(* IEC 61131-3 sources: daoli-st-library/DL_Process (part 34) *)

(* ---- FB_DL_FirstArticleLock.st ---- *)
(*
  ==================================================================
  组件名 Component  : FB_DL_FirstArticleLock
  分类   Category   : DL_Process
  复杂度 Complexity  : cx5
  版本   Version    : 1.0.0
  功能   Purpose    : 首件检验锁定。首件未放行禁止批量运行（许可出口挂锁定
                      状态量）；换型信号沿自动重锁；首件检验合格沿解锁放行
                      并出单拍放行脉冲与台账；锁定期的运行请求出单拍拒绝
                      指示。汽车 / 电子行业公开首件流程语义。
  来源   Source     : self（行业公开流程）
  溯源   Origin     : IEC 61131-3 标准语义的道莅防御性实现；首件检验锁定为
                      公开行业流程语义，clean-room 自研实现，未复制任何厂商
                      私有库源码。
  平台   Platform   : 纯 IEC 61131-3（Standard.library: R_TRIG，无私有库）
  分工声明 Split     : 与 FB_DL_MaterialHoldTimeEnforce 分工——保持时限件做
                      在制批次时限门控，本件做换型后批量运行前置门控；与
                      存量批次追溯件分工——本件不含履历数据，只有锁存与台账。
  作者   Author     : 道莅代码库 · PLC 编程专家（R58）
  ------------------------------------------------------------------
  边界 Boundary     :
                      一 上电默认锁定（_bInit 首扫置锁）：首件未放行禁止批
                         量运行，安全侧缺省；
                      二 锁定解除路径 = bFaPass 上升沿（唯一解锁路径，R188
                         头注释声明）；重锁路径 = bChangeover 上升沿（换型
                         自动重锁）；
                      三 许可出口挂状态量 _bLocked（R99：禁挂单拍标志）；
                      四 单拍标志 bFaRelease / bRunBlocked 每拍预清零（R25，
                         置位点在段 3，统一出口单拍映射两段式 R189）；
                      五 复位沿作用域：清台账 / 恢复默认锁定（两项逐项声明）；
                      六 无全局变量、无外部变量声明、无物理地址寻址。
  修订记录 Revision  :
    2026-11-21  v1.0.0  R58 首版（批 4 · 序号 16）
  ==================================================================
*)

FUNCTION_BLOCK FB_DL_FirstArticleLock
VAR_INPUT
    bEnable     : BOOL := TRUE;   // 使能，失能许可出口安全侧 FALSE [-] / enable, disabling clears the permit
    bReset      : BOOL := FALSE;  // 复位上升沿清台账并恢复默认锁定 [-] / reset rising edge clears the ledger and restores the default lock
    bChangeover : BOOL := FALSE;  // 换型信号（沿生效，自动重锁）[-] / the changeover signal, edge effective, auto relock
    bFaPass     : BOOL := FALSE;  // 首件检验合格（沿生效）[-] / the first article pass, edge effective
    bRunReq     : BOOL := FALSE;  // 批量运行请求电平 [-] / the batch run request level
END_VAR
VAR_OUTPUT
    bBatchPermit: BOOL := FALSE; // 批量运行许可出口（挂锁定状态量）[-] / the batch run permit outlet, gated by the lock state
    bLocked     : BOOL := FALSE; // 锁定中指示出口 [-] / the locked indicator outlet
    bFaRelease  : BOOL := FALSE; // 首件放行单拍出口 [-] / the first article release pulse outlet
    bRunBlocked : BOOL := FALSE; // 锁定期运行请求拒绝单拍出口 [-] / the run request blocked pulse outlet
    nLockCnt    : UDINT := 0;    // 累计重锁次数 [次] / the total relock count
    nRelCnt     : UDINT := 0;    // 累计放行次数 [次] / the total release count
END_VAR
VAR
    rtChg   : R_TRIG; // 换型沿检测，段 0 无条件刷新 / the changeover edge
    rtPass  : R_TRIG; // 首件合格沿检测，段 0 无条件刷新 / the pass edge
    rtReset : R_TRIG; // 复位沿检测，段 0 无条件刷新 / the reset edge
    _bLocked: BOOL := TRUE;  // 锁定状态量（上电缺省锁定，边界一）/ the lock state, the power up default locked
    _bRel   : BOOL := FALSE; // 放行脉冲内部保持量（统一出口映射单拍）/ the release pulse internal holder
    _bBlk   : BOOL := FALSE; // 拒绝脉冲内部保持量 / the blocked pulse internal holder
    _bInit  : BOOL := FALSE; // 首扫初始化完成标志（R310）/ the first scan flag
END_VAR
VAR CONSTANT
    DL_FAL_CNTMAX : UDINT := 4294967294; // 台账计数钳定界 [次]，防 UDINT 回绕 / the ledger clamp against a wrap
END_VAR

// 段 0｜沿检测无条件周期刷新（禁入分支，FB50-1）/ segment 0, the unconditional refresh
rtChg(CLK := bChangeover); // 换型沿 / the changeover edge
rtPass(CLK := bFaPass); // 合格沿 / the pass edge
rtReset(CLK := bReset); // 复位沿 / the reset edge

// 段 1｜首扫初始化（R310）：上电默认锁定（边界一）/ segment 1, the first scan, the default locked
IF NOT _bInit THEN // 首扫一拍 / the first scan
    _bInit := TRUE; // 置首扫标志 / raise the flag
    _bLocked := TRUE; // 上电默认锁定 / the default locked
END_IF

// 段 2｜复位沿作用域：清台账 / 恢复默认锁定（两项逐项声明，边界五）/ segment 2, the reset edge scope
IF rtReset.Q THEN // 复位沿 / the reset edge
    nLockCnt := 0; // 作用域一：清重锁台账 / scope one, clear the relock ledger
    nRelCnt := 0; // 作用域一：清放行台账 / scope one, clear the release ledger
    _bLocked := TRUE; // 作用域二：恢复默认锁定（安全侧）/ scope two, restore the default lock
END_IF

// 段 3｜重锁与解锁沿判定 + 单拍保持量置位（边界二三四）/ segment 3, the relock and the unlock edges
IF rtChg.Q THEN // 换型沿自动重锁 / the changeover edge relocks
    _bLocked := TRUE; // 置锁定 / raise the lock
    IF nLockCnt < DL_FAL_CNTMAX THEN // 台账防回绕 / the ledger wrap guard
        nLockCnt := nLockCnt + 1; // 重锁台账推进 / advance the relock ledger
    END_IF
END_IF
IF _bLocked AND rtPass.Q THEN // 锁定中且首件合格沿（唯一解锁路径，R188）/ locked with the pass edge
    _bLocked := FALSE; // 解锁 / release the lock
    IF nRelCnt < DL_FAL_CNTMAX THEN // 台账防回绕 / the ledger wrap guard
        nRelCnt := nRelCnt + 1; // 放行台账推进 / advance the release ledger
    END_IF
    _bRel := TRUE; // 置放行内部保持量 / raise the release holder
END_IF
IF _bLocked AND bRunReq THEN // 锁定期收到运行请求 / a run request while locked
    _bBlk := TRUE; // 置拒绝内部保持量 / raise the blocked holder
END_IF
bFaRelease := FALSE; // 放行单拍每拍预清零（R25）/ the release pulse preset false each scan
bRunBlocked := FALSE; // 拒绝单拍每拍预清零（R25）/ the blocked pulse preset false each scan

// 段 4｜统一出口（边界三四：状态量门控 + 单拍两段式映射）/ segment 4, the unified outlet
bBatchPermit := (NOT _bLocked) AND bEnable; // 许可挂锁定状态量（R99）/ the permit gated by the lock state
bLocked := _bLocked; // 锁定指示同源 / the indicator shares the state
IF _bRel THEN // 放行保持量 → 统一出口单拍映射（两段式，R189）/ the holder mapped to the pulse
    bFaRelease := TRUE; // 放行单拍 / the release pulse
    _bRel := FALSE; // 消费保持量 / consume the holder
END_IF
IF _bBlk THEN // 拒绝保持量 → 统一出口单拍映射 / the holder mapped to the pulse
    bRunBlocked := TRUE; // 拒绝单拍 / the blocked pulse
    _bBlk := FALSE; // 消费保持量 / consume the holder
END_IF
END_FUNCTION_BLOCK

(* ---- FB_DL_FloatBathTopRollSeq.st ---- *)
(*
  Name: FB_DL_FloatBathTopRollSeq
  Category: DL_Process
  Version: 1.0.0
  Round: R90 / 2026-11-25
  开源溯源：clean-room 自研（族 浮法玻璃锡槽退火，ST 开源生态实测 0 命中，无外部代码引入）
  功能：1) 拉边机三轴同步作业序，六相推进：待机 → 就位 → 夹持 → 同步张角 → 跟踪带宽 → 退出 → 完成。
           就位相向三轴发出就位指令并等三路到位信号全为 TRUE；夹持相保持指令并等夹持时长；
           同步张角相把张角给定按设定角速度斜坡推到 fAngleTargetDeg；跟踪带宽相保持张角并监视
           带宽是否漂出容差；退出相撤令（三轴回退），等退到位时长后置完成位。
        2) 多轴失步监视贯穿三轴：就位相超时未全部到位 → 失步故障；同步相与跟踪相内任一路到位
           信号掉线 → 失步故障。三轴指令始终同源（同一个状态量导出），不存在单轴独走的可能。
        3) 张角斜坡按「角速度 × 扫描周期」逐拍累加，故扫描周期必须作为入参并做零闸（R21），
           不许假设固定扫描周期；斜坡单向逼近目标，不越过目标值。
  边界条件：1) 非有限值闸：张角目标、带宽实测、扫描周期三路实值入参统一过
           NOT(x > -DL_BIG AND x < DL_BIG)，同时拦 NaN 与 Inf；命中即判组态非法并进故障相，
           绝不把 NaN 累加进张角保持值（累加后保持值被永久污染，R19）。
        2) 组态零闸：ABS(fCycleS) > DL_EPS 才允许角度积分（周期为零则斜坡不推进且步进发散）；
           tSyncS 必须 > T#0S（跟踪相时长为 0 表示跳过跟踪监视，属组态错误）；
           fAngleTargetDeg 必须落在 0 ~ DL_ANGLE_MAX_DEG(90 °) 并大于 0。
        3) 带宽容差闸：跟踪相内带宽相对漂移超过 DL_WIDTH_TOL_PCT(2 %) 判带宽失控故障；
           带宽参考值在进入跟踪相的同一个周期末锁存（R23：快照必须在迁移判断之后更新）。
        4) 相超时说明：eFbtPosition 由 tonPos 监视（就位超时 = 失步）；
           eFbtClamp 由 tonClamp 定时（夹持时长，无额外超时）；
           eFbtSyncAngle 由 tonAngle 监视（张角同步超时 = 失步）；
           eFbtTrackWidth 由 tonTrack 定时（跟踪时长，另有带宽容差监视）；
           eFbtRetract 由 tonRetract 定时（退出时长）；
           eFbtDone / eFbtIdle / eFbtFault 为稳态持留相，不设相超时（设了会周期性误报）；
           整序另设 tonSeq 总超时兜底。
        5) 状态机兜底：CASE 全态覆盖 + ELSE 强制回故障相并撤全部指令；故障解除路径为
           (NOT xStart) AND (NOT xFault) AND 组态恢复，可达。
        6) FB 主体不使用 RETURN，统一单出口（跨平台可移植性）。
  量纲自证：张角步进 = (°/s) × s = °，与 fAngleDeg 同量纲；
           带宽相对漂移 = (mm − mm) / mm × 100 = 无因次 [%]，与容差同量纲；
           三路到位信号为 [bool]；tonXxx 的 PT 均为 [TIME]；本件无跨量纲相加。
  码表 Error codes（本件格 0090_07xx，故障级一律 3 行内置 _uFault/_bFault/_eState）:
    16#0090_0701 故障级：组态非法（角度目标/跟踪时长/扫描周期越界或非有限）
    16#0090_0702 故障级：就位超时（三轴未全部到位，多轴失步）
    16#0090_0703 故障级：张角同步超时（斜坡未在时限内到达目标）
    16#0090_0704 故障级：同步/跟踪相内到位信号掉线（多轴失步）
    16#0090_0705 故障级：跟踪相带宽漂移超容差（带宽失控）
    16#0090_0706 故障级：整序总超时
    16#0090_0707 故障级：外部故障输入 xFault
    16#0090_0708 故障级：状态机落 ELSE 兜底（非法相位 ID）
    16#0090_0709 信息级：张角已到达目标，转入跟踪相

  修订历史 Revision :
    2026-11-25  v1.0.0  R90 首版
*)

TYPE E_DL_FbtState :
(
    eFbtIdle      := 0,    // 待机：等启动上升沿 / Idle, awaiting start edge
    eFbtPosition  := 10,   // 就位：三轴发出就位指令 / Positioning, all three axes commanded
    eFbtClamp     := 20,   // 夹持：保持指令等夹持时长 / Clamping, commands held
    eFbtSyncAngle := 30,   // 同步张角：斜坡推到目标角 / Angle synchronising
    eFbtTrackWidth:= 40,   // 跟踪带宽：保持张角并监视带宽 / Width tracking
    eFbtRetract   := 50,   // 退出：撤令等退到位 / Retracting
    eFbtDone      := 60,   // 完成：保持完成位等撤令 / Done, held until release
    eFbtFault     := 90    // 故障：锁存待解除 / Fault, latched awaiting release
);
END_TYPE

FUNCTION_BLOCK FB_DL_FloatBathTopRollSeq
VAR_INPUT
    xStart          : BOOL;    // 作业启动指令（上升沿有效）[bool] / Sequence start, edge triggered [bool]
    xFault          : BOOL;    // 外部故障汇总 [bool] / External fault aggregate [bool]
    xInPos1         : BOOL;    // 1 轴到位信号 [bool] / Axis 1 in-position signal [bool]
    xInPos2         : BOOL;    // 2 轴到位信号 [bool] / Axis 2 in-position signal [bool]
    xInPos3         : BOOL;    // 3 轴到位信号 [bool] / Axis 3 in-position signal [bool]
    fAngleTargetDeg : REAL;    // 目标张角 [°] / Target nip angle [°]
    fWidthMeasMm    : REAL;    // 玻璃带宽度实测 [mm] / Measured ribbon width [mm]
    tSyncS          : TIME;    // 带宽跟踪监视时长 [TIME] / Width tracking supervision duration [TIME]
    fCycleS         : REAL;    // 扫描周期 [s] / Scan cycle time [s]
END_VAR
VAR_OUTPUT
    xCmd1           : BOOL;    // 1 轴就位/夹持指令 [bool] / Axis 1 command [bool]
    xCmd2           : BOOL;    // 2 轴就位/夹持指令 [bool] / Axis 2 command [bool]
    xCmd3           : BOOL;    // 3 轴就位/夹持指令 [bool] / Axis 3 command [bool]
    fAngleDeg       : REAL;    // 当前张角给定 [°] / Current nip angle setpoint [°]
    fWidthDevPct    : REAL;    // 跟踪相带宽相对漂移 [%] / Width relative drift during tracking [%]
    xAllInPos       : BOOL;    // 三轴全部到位 [bool] / All three axes in position [bool]
    xDone           : BOOL;    // 作业完成保持位 [bool] / Sequence complete held flag [bool]
    eState          : E_DL_FbtState;   // 状态出口，段尾单点映射 / State outlet, single-point mapped
    nErrId          : UDINT;   // 事件码，0 = 无事件 / Event code, 0 = none
END_VAR
VAR
    tonPos          : TON;     // 就位相超时监视 [TIME] / Positioning timeout timer
    tonClamp        : TON;     // 夹持时长定时 [TIME] / Clamping duration timer
    tonAngle        : TON;     // 张角同步超时监视 [TIME] / Angle synchronising timeout timer
    tonTrack        : TON;     // 带宽跟踪时长定时 [TIME] / Width tracking duration timer
    tonRetract      : TON;     // 退出相时长定时 [TIME] / Retracting duration timer
    tonSeq          : TON;     // 整序总超时定时 [TIME] / Whole-sequence timeout timer
    rtStart         : R_TRIG;  // 启动上升沿检测 [bool] / Start rising edge detector
    _eState         : E_DL_FbtState := E_DL_FbtState.eFbtIdle;   // 内部相位（CASE 唯一写入目标）
    _eStatePrev     : E_DL_FbtState := E_DL_FbtState.eFbtIdle;   // 上一拍相位快照（周期末更新）
    _fAngleDeg      : REAL;    // 张角保持值 [°] / Retained nip angle [°]
    _fWidthRefMm    : REAL;    // 跟踪相带宽参考值（进相锁存）[mm] / Width reference latched on entry [mm]
    _fWidthDevPct   : REAL;    // 带宽相对漂移 [%] / Width relative drift [%]
    _fStepDeg       : REAL;    // 单拍张角步进 [°] / Angle step per cycle [°]
    _bAllInPos      : BOOL;    // 三轴全到位 [bool] / All axes in position [bool]
    _bCmdOut        : BOOL;    // 三轴指令聚合（状态导出）[bool] / Axis command aggregate [bool]
    _bCfgBad        : BOOL;    // 组态非法聚合 [bool] / Configuration invalid aggregate [bool]
    _bActive        : BOOL;    // 序激活（中间五相）[bool] / Sequence active flag [bool]
    _bAngleAtTgt    : BOOL;    // 张角已到目标（带死区）[bool] / Angle reached target [bool]
    _bWidthBad      : BOOL;    // 带宽漂移超容差 [bool] / Width drift out of tolerance [bool]
    _bFault         : BOOL;    // 故障锁存位 [bool] / Latched fault flag [bool]
    _uInfo          : UDINT;   // 信息码，每拍重算 / Info code, recomputed every cycle
    _uFault         : UDINT;   // 故障码锁存 / Latched fault code
END_VAR
VAR CONSTANT
    DL_EPS          : REAL := 1.0E-9;    // 组态零闸阈值 [-] / Configuration zero gate threshold [-]
    DL_BIG          : REAL := 1.0E12;    // 非有限值闸量级上限 [-] / Finiteness gate magnitude [-]
    DL_PCT          : REAL := 100.0;     // 百分比换算因子 [%] / Percent conversion factor [%]
    DL_ANGLE_MAX_DEG: REAL := 90.0;      // 张角量程上限 [°] / Nip angle range ceiling [°]
    DL_ANGLE_RATE   : REAL := 2.0;       // 张角斜坡角速度 [°/s] / Angle ramp rate [°/s]
    DL_ANGLE_TOL_DEG: REAL := 0.10;      // 张角到位死区 [°] / Angle arrival deadband [°]
    DL_WIDTH_TOL_PCT: REAL := 2.0;       // 带宽漂移容差 [%] / Width drift tolerance [%]
    DL_POS_MAX      : TIME := T#20S;     // 就位相超时上限 [TIME] / Positioning timeout ceiling [TIME]
    DL_CLAMP_S      : TIME := T#3S;      // 夹持时长 [TIME] / Clamping duration [TIME]
    DL_ANGLE_MAX_T  : TIME := T#60S;     // 张角同步超时上限 [TIME] / Angle timeout ceiling [TIME]
    DL_RETRACT_S    : TIME := T#8S;      // 退出相时长 [TIME] / Retracting duration [TIME]
    DL_SEQ_MAX      : TIME := T#15M;     // 整序总超时上限 [TIME] / Whole-sequence timeout [TIME]
END_VAR

(* —— 段 0：单拍量预清零（锁存量 _uFault/_bFault/_fAngleDeg/_fWidthRefMm/_eStatePrev 不入清单） —— *)
_uInfo := 16#0000_0000;                     // 信息码每拍重算 / Info code recomputed
nErrId := 16#0000_0000;                     // 事件码缺省无事件 / Event code defaults to none
_fWidthDevPct := 0.0;                       // 带宽漂移每拍重算 / Width drift recomputed

(* —— 段 1：非有限值闸（R19：NaN 一旦累加进保持值会永久污染，必须前置拦截） —— *)
_bCfgBad := NOT (fAngleTargetDeg > -DL_BIG AND fAngleTargetDeg < DL_BIG)
            OR NOT (fWidthMeasMm > -DL_BIG AND fWidthMeasMm < DL_BIG)
            OR NOT (fCycleS > -DL_BIG AND fCycleS < DL_BIG);

(* —— 段 2：组态零闸（R4 / R21：周期零闸是角度积分的前置条件） —— *)
_bCfgBad := _bCfgBad
            OR (ABS(fCycleS) <= DL_EPS)                      // 周期为零：角度积分不推进且发散
            OR (tSyncS <= T#0S)                              // 跟踪时长为零：跳过监视属错组态
            OR (fAngleTargetDeg <= DL_EPS)                   // 目标张角必须为正
            OR (fAngleTargetDeg > DL_ANGLE_MAX_DEG);         // 目标张角不得越量程

(* —— 段 3：状态派生与判据量 —— *)
_fStepDeg := LIMIT(0.0, DL_ANGLE_RATE * fCycleS, DL_ANGLE_MAX_DEG);   // °/s × s = °
_bAllInPos := xInPos1 AND xInPos2 AND xInPos3;                        // 三轴全到位
_bAngleAtTgt := (NOT _bCfgBad) AND (ABS(fAngleTargetDeg - _fAngleDeg) <= DL_ANGLE_TOL_DEG);
_bActive := (_eState = E_DL_FbtState.eFbtPosition) OR (_eState = E_DL_FbtState.eFbtClamp)
            OR (_eState = E_DL_FbtState.eFbtSyncAngle) OR (_eState = E_DL_FbtState.eFbtTrackWidth)
            OR (_eState = E_DL_FbtState.eFbtRetract);
_bCmdOut := (_eState = E_DL_FbtState.eFbtPosition) OR (_eState = E_DL_FbtState.eFbtClamp)
            OR (_eState = E_DL_FbtState.eFbtSyncAngle) OR (_eState = E_DL_FbtState.eFbtTrackWidth);

(* 带宽相对漂移：分母零闸后才允许相除（参考值在跟踪相入口锁存） *)
IF ABS(_fWidthRefMm) > DL_EPS THEN
    _fWidthDevPct := (fWidthMeasMm - _fWidthRefMm) / _fWidthRefMm * DL_PCT;   // [%]
ELSE
    _fWidthDevPct := 0.0;                                                 // 参考值不可用则不计漂移
END_IF
_bWidthBad := (_eState = E_DL_FbtState.eFbtTrackWidth) AND (ABS(_fWidthDevPct) > DL_WIDTH_TOL_PCT);

(* —— 段 4：定时器与边沿无条件周期刷新（R7：调用语句不得置于 IF/CASE 内） —— *)
rtStart(CLK := xStart);                                                             // 启动上升沿
tonPos(IN := (_eState = E_DL_FbtState.eFbtPosition), PT := DL_POS_MAX);             // 就位超时监视
tonClamp(IN := (_eState = E_DL_FbtState.eFbtClamp), PT := DL_CLAMP_S);              // 夹持时长
tonAngle(IN := (_eState = E_DL_FbtState.eFbtSyncAngle), PT := DL_ANGLE_MAX_T);      // 张角同步超时
tonTrack(IN := (_eState = E_DL_FbtState.eFbtTrackWidth), PT := tSyncS);             // 跟踪时长
tonRetract(IN := (_eState = E_DL_FbtState.eFbtRetract), PT := DL_RETRACT_S);        // 退出时长
tonSeq(IN := _bActive, PT := DL_SEQ_MAX);                                           // 整序总超时

(* —— 段 5：全局故障拦截（优先级最高；已锁存则不再改写码值，禁同拍抹除） —— *)
IF xFault AND (NOT _bFault) THEN
    _uFault := 16#0090_0707;                // 故障级：外部故障输入
    _bFault := TRUE;                        // 锁存（3 行内置，R45 配对）
    _eState := E_DL_FbtState.eFbtFault;
END_IF
IF _bCfgBad AND (NOT _bFault) THEN
    _uFault := 16#0090_0701;                // 故障级：组态非法
    _bFault := TRUE;                        // 锁存
    _eState := E_DL_FbtState.eFbtFault;
END_IF
IF tonSeq.Q AND _bActive AND (NOT _bFault) THEN
    _uFault := 16#0090_0706;                // 故障级：整序总超时
    _bFault := TRUE;                        // 锁存
    _eState := E_DL_FbtState.eFbtFault;
END_IF
IF _bWidthBad AND (NOT _bFault) THEN
    _uFault := 16#0090_0705;                // 故障级：跟踪相带宽漂移超容差
    _bFault := TRUE;                        // 锁存
    _eState := E_DL_FbtState.eFbtFault;
END_IF

(* —— 段 6：相位机（只做迁移；出口在段 8 单点映射） —— *)
CASE _eState OF

E_DL_FbtState.eFbtIdle:
    IF NOT xStart THEN
        ;                                   // 等启动 / Waiting for start
    ELSIF rtStart.Q THEN
        _eState := E_DL_FbtState.eFbtPosition;   // 进就位相
    END_IF

E_DL_FbtState.eFbtPosition:
    IF NOT xStart THEN
        _eState := E_DL_FbtState.eFbtIdle;      // 撤令：回待机
    ELSIF _bAllInPos THEN
        _eState := E_DL_FbtState.eFbtClamp;     // 三轴全到位：进夹持相
    ELSIF tonPos.Q THEN
        _uFault := 16#0090_0702;                // 故障级：就位超时（多轴失步）
        _bFault := TRUE;
        _eState := E_DL_FbtState.eFbtFault;
    END_IF

E_DL_FbtState.eFbtClamp:
    IF NOT xStart THEN
        _eState := E_DL_FbtState.eFbtIdle;
    ELSIF NOT _bAllInPos THEN
        _uFault := 16#0090_0704;                // 故障级：夹持中到位信号掉线（多轴失步）
        _bFault := TRUE;
        _eState := E_DL_FbtState.eFbtFault;
    ELSIF tonClamp.Q THEN
        _eState := E_DL_FbtState.eFbtSyncAngle; // 夹持完成：进同步张角相
    END_IF

E_DL_FbtState.eFbtSyncAngle:
    IF NOT xStart THEN
        _eState := E_DL_FbtState.eFbtIdle;
    ELSIF NOT _bAllInPos THEN
        _uFault := 16#0090_0704;                // 故障级：同步中到位信号掉线（多轴失步）
        _bFault := TRUE;
        _eState := E_DL_FbtState.eFbtFault;
    ELSIF _bAngleAtTgt THEN
        _uInfo := 16#0090_0709;                 // 信息级：张角已到达目标
        _eState := E_DL_FbtState.eFbtTrackWidth; // 本拍合法事件优先于超时迁移（R275）
    ELSIF tonAngle.Q THEN
        _uFault := 16#0090_0703;                // 故障级：张角同步超时
        _bFault := TRUE;
        _eState := E_DL_FbtState.eFbtFault;
    ELSE
        _fAngleDeg := MIN(fAngleTargetDeg, _fAngleDeg + _fStepDeg);   // 单向逼近，不越目标
    END_IF

E_DL_FbtState.eFbtTrackWidth:
    IF NOT xStart THEN
        _eState := E_DL_FbtState.eFbtIdle;
    ELSIF NOT _bAllInPos THEN
        _uFault := 16#0090_0704;                // 故障级：跟踪中到位信号掉线（多轴失步）
        _bFault := TRUE;
        _eState := E_DL_FbtState.eFbtFault;
    ELSIF tonTrack.Q THEN
        _eState := E_DL_FbtState.eFbtRetract;   // 跟踪结束：进退出相
    END_IF

E_DL_FbtState.eFbtRetract:
    IF xFault THEN
        _uFault := 16#0090_0707;                // 故障级：退出中外部故障
        _bFault := TRUE;
        _eState := E_DL_FbtState.eFbtFault;
    ELSIF tonRetract.Q THEN
        _eState := E_DL_FbtState.eFbtDone;      // 退到位：进完成相
    END_IF

E_DL_FbtState.eFbtDone:
    IF NOT xStart THEN
        _eState := E_DL_FbtState.eFbtIdle;      // 撤令：回待机
    END_IF

E_DL_FbtState.eFbtFault:
    IF (NOT xStart) AND (NOT xFault) AND (NOT _bCfgBad) THEN
        _bFault := FALSE;                       // 解除路径：撤令 + 外部故障消失 + 组态恢复（可达）
        _uFault := 16#0000_0000;                // 清锁存码
        _eState := E_DL_FbtState.eFbtIdle;      // 回待机
    END_IF

ELSE
    _uFault := 16#0090_0708;                    // 故障级：非法相位 ID 兜底
    _bFault := TRUE;                            // 锁存
    _eState := E_DL_FbtState.eFbtFault;         // 强制回故障相

END_CASE

(* —— 段 7：后置段（R23：带宽参考快照在迁移判断之后按「进入沿」锁存） —— *)
IF (_eState = E_DL_FbtState.eFbtTrackWidth) AND (_eStatePrev <> E_DL_FbtState.eFbtTrackWidth) THEN
    _fWidthRefMm := fWidthMeasMm;               // 进跟踪相当拍锁存带宽参考值 [mm]
END_IF
IF _eState <> E_DL_FbtState.eFbtTrackWidth THEN
    _fWidthRefMm := fWidthMeasMm;               // 非跟踪相：参考值持续跟随，避免陈旧值误判
END_IF
_eStatePrev := _eState;                         // 快照统一在周期末尾更新（R23）

(* —— 段 8：出口单点映射（名实同源；三轴指令同源导出，故障侧一律撤令） —— *)
xCmd1 := _bCmdOut AND (NOT _bFault);            // 1 轴指令出口
xCmd2 := _bCmdOut AND (NOT _bFault);            // 2 轴指令出口
xCmd3 := _bCmdOut AND (NOT _bFault);            // 3 轴指令出口
fAngleDeg := LIMIT(0.0, _fAngleDeg, DL_ANGLE_MAX_DEG);   // 张角给定出口 [°]
fWidthDevPct := LIMIT(-DL_BIG, _fWidthDevPct, DL_BIG);   // 带宽漂移出口 [%]
xAllInPos := _bAllInPos;                                 // 三轴到位出口
xDone := (_eState = E_DL_FbtState.eFbtDone) AND (NOT _bFault);   // 完成位出口
eState := _eState;                                       // 状态出口单点映射
IF _bFault THEN
    nErrId := _uFault;                          // 故障锁存码回放（不在故障相按当下输入重推断）
ELSE
    nErrId := _uInfo;                           // 信息码
END_IF

END_FUNCTION_BLOCK

(* ---- FB_DL_FlowTotalizer.st ---- *)
(*==============================================================================
 * 组件名称 (Component)  : FB_DL_FlowTotalizer
 * 所属子库 (Sublibrary) : DL_Process
 * 前缀     (Prefix)     : FB_DL_
 * 当前版本 (Version)    : 1.0.0
 * 兼容性   (Platform)   : CODESYS 3.5 / TwinCAT 3 / 汇川 InoProShop / Schneider
 *                         Machine Expert；纯 IEC 61131-3（第 3 版），
 *                         仅依赖标准库 TON / R_TRIG / ABS / MAX / MIN，零厂商方言
 * 作者     (Author)     : 道莅代码库 · PLC编程专家（R31）
 * 开源溯源 (Origin)     : 流量累积与批控公开语义（行业池），道莅 clean-room
 *                         防御性实现，未复制任何外部源码行
 * 功能描述 (Function)   : 流量累积与批控零点件。累积量 ΔV = fFlow·Δt，Δt 取
 *                         实际运行时间差（计时器实测经过值差分，非定时器
 *                         假设值）防扫描抖动误差；清零沿先保存结算快照再
 *                         清批次；寿命累计饱和于 DL_TOTAL_MAX 防溢出。
 *                         与库内 EnergyMeterAccum 边界：该件为千瓦时电量
 *                         口径，本件为升流量口径，二者不合并。
 * 码位     (Codes)      : 16#0005_00AD 信息级：流量非有限按零积分、Δt 越界
 *                                      按上次有效值钳位、批满提示（不置
 *                                      bError，规格仅信息级）
 *                         16#0005_00AE~00B1 保留未启用（码表与实现对齐）
 *                         偏离：uErrorId 规格标 UINT，段位码超 UINT 值域，
 *                         按 32 位载体 UDINT 落地（与库内段位码惯例一致）
 * 边界防错 (Boundary)   : 1 fFlow 非有限本拍按 0 积分记信息码不中断；
 *                         2 Δt 不大于零或超扫描周期 10 倍按上次有效值钳位；
 *                         3 清零沿与积分同拍冲突先积分后清零（不丢该拍）；
 *                         4 bBatchFull 置位有销位路径：bRstBatch 清零沿；
 *                         5 TON/R_TRIG 实例每拍无条件刷新；
 *                         6 首扫同步时标基准防上电尖峰。
 * 修订历史 (Revision)   : 2026-11-18 v1.0.0 首版入库（R31 · 阶段三 · 序 15）
 *==============================================================================*)

(*==============================================================================
 * 功能块: FB_DL_FlowTotalizer
 * 调用约定: 每个扫描周期无条件调用一次；tSample 为名义采样周期（钳位判据
 *           用），实际 Δt 取计时器经过值差分。
 *==============================================================================*)
FUNCTION_BLOCK FB_DL_FlowTotalizer
VAR_INPUT
    fFlow      : REAL := 0.0;         // 瞬时流量 [升每分钟] / Instantaneous flow [L per min]
    bRstBatch  : BOOL := FALSE;        // 批次清零沿 / Batch reset edge
    bEn        : BOOL := FALSE;        // 使能 / Enable flag
    tSample    : TIME := T#1S;         // 名义采样周期 [毫秒]（钳位判据基准）/ Nominal sample period [ms], clamp basis
    fBatchLimit: REAL := 1000.0;      // 批量限值 [升]（可增引脚）/ Batch volume limit [L], added pin
END_VAR
VAR_OUTPUT
    fTotalBatch: REAL;                 // 批次累计量 [升] / Batch total [L]
    fTotalLife : REAL;                 // 寿命累计量 [升] / Lifetime total [L]
    bBatchFull : BOOL;                 // 批满标志（清零沿销位）/ Batch full flag, cleared by reset edge
    uErrorId   : UDINT;                // 信息级码，0 = 无信息（段位码 32 位载体，规格 UINT 值域不足，偏离留档）/ Info code, 0 = none, 32-bit carrier deviation
END_VAR
VAR
    rTrigRst   : R_TRIG;               // 清零沿检测，每拍无条件刷新 / Reset edge detector, refreshed every scan
    tonMeter   : TON;                  // 实际运行时标（大超时经过值表）/ Run-time meter, elapsed register
    fEtPrev    : REAL;                 // 上拍经过值 [毫秒] / Previous elapsed [ms]
    fEtNow     : REAL;                 // 本拍经过值 [毫秒] / Current elapsed [ms]
    fDtMs      : REAL;                 // 有效时间差 [毫秒] / Effective delta time [ms]
    fDtSec     : REAL;                 // 有效时间差 [秒] / Effective delta time [s]
    bFirst     : BOOL := TRUE;         // 首扫标志 / First-scan flag
    fBatchSnap : REAL;                 // 清零前结算快照 [升] / Batch snapshot before reset [L]
    bFlowBad   : BOOL;                 // 本拍流量非有限 / Flow non-finite this scan
    bDtClamp   : BOOL;                 // 本拍 Δt 越界钳位 / Delta time clamped this scan
    fFlowEff   : REAL;                 // 本拍生效流量 [升每分钟] / Effective flow [L per min]
END_VAR
VAR CONSTANT
    DL_FT_FIN     : REAL  := 1.0E30;   // REAL 有限幅值判界 / REAL finiteness magnitude bound
    DL_FT_DTMAXF  : REAL  := 10.0;     // Δt 越界倍率（名义周期十倍）/ Delta time overrange factor
    DL_FT_TOTALMAX: REAL  := 1.0E12;   // 寿命累计饱和上限 [升] / Lifetime saturation ceiling [L]
    DL_FT_SEC     : REAL  := 1000.0;   // 毫秒到秒换算系数 / Millisecond to second factor
END_VAR

// ---- 段 1｜边沿与计时实例无条件刷新（红线：禁入条件分支）----------------------
rTrigRst(CLK := bRstBatch);                           // 清零沿检测 / Reset edge detection
tonMeter(IN := bEn, PT := T#4294967MS);               // 运行时标，使能即累计 / Run-time meter, accumulates while enabled

// ---- 段 2｜实际时间差分（非定时器假设值）--------------------------------------
fEtNow := TIME_TO_REAL(tonMeter.ET);                  // 本拍经过值 [毫秒] / Current elapsed [ms]
fDtMs  := fEtNow - fEtPrev;                           // 实际时间差 [毫秒] / Real delta time [ms]
bDtClamp := FALSE;                                    // 钳位标志先清 / Clear clamp flag
IF bFirst OR (fDtMs <= 0.0) OR (fDtMs > TIME_TO_REAL(tSample) * DL_FT_DTMAXF) THEN
    fDtMs := TIME_TO_REAL(tSample);                   // 首扫或越界按名义周期钳位 / First scan or out-of-range clamped
    bDtClamp := NOT bFirst;                           // 非首扫才记钳位信息 / Clamp info only after first scan
END_IF
fEtPrev := fEtNow;                                    // 快照留痕 / Snapshot previous elapsed
bFirst := FALSE;                                      // 清首扫标志 / Clear first-scan flag
fDtSec := fDtMs / DL_FT_SEC;                          // 换算秒 [秒] / Convert to seconds

// ---- 段 3｜流量有效性（非有限按零积分不中断）----------------------------------
bFlowBad := (fFlow <> fFlow) OR (ABS(fFlow) >= DL_FT_FIN); // 流量非有限判定 / Flow non-finite detection
IF bFlowBad THEN
    fFlowEff := 0.0;                                  // 非有限按零积分 / Non-finite integrates as zero
ELSE
    fFlowEff := fFlow;                                // 有效原值 / Valid value as-is
END_IF

// ---- 段 4｜积分（先积分后清零：同拍冲突不丢该拍）------------------------------
IF bEn THEN
    fTotalBatch := fTotalBatch + fFlowEff * fDtSec / 60.0; // 批次积分 ΔV=f·Δt / Batch integrates flow over time
    IF fTotalLife < DL_FT_TOTALMAX THEN
        fTotalLife := MIN(fTotalLife + fFlowEff * fDtSec / 60.0, DL_FT_TOTALMAX); // 寿命累计饱和防溢出 / Lifetime saturates
    END_IF
END_IF

// ---- 段 5｜批满判定（置位有销位路径：清零沿）----------------------------------
IF fTotalBatch >= fBatchLimit THEN
    bBatchFull := TRUE;                               // 批满置位 / Batch full set
END_IF

// ---- 段 6｜清零沿：先保存结算快照再清批次（批满标志同拍销位）------------------
IF rTrigRst.Q THEN
    fBatchSnap  := fTotalBatch;                       // 结算快照留档 / Settlement snapshot kept
    fTotalBatch := 0.0;                               // 批次清零 / Batch cleared
    bBatchFull  := FALSE;                             // 批满标志销位 / Batch full cleared
END_IF

// ---- 段 7｜信息级码装配（不置故障标志，规格仅信息级）--------------------------
IF bFlowBad OR bDtClamp THEN
    uErrorId := 16#0005_00AD;                         // 信息级：非有限/钳位 / Info: non-finite or clamp
ELSIF bBatchFull THEN
    uErrorId := 16#0005_00AD;                         // 信息级：批满提示 / Info: batch full
ELSE
    uErrorId := 16#0000_0000;                         // 无码 / No code
END_IF
END_FUNCTION_BLOCK

(* ---- FB_DL_ForelinePressureCtrl.st ---- *)
(*
  FB_DL_ForelinePressureCtrl  —  真空前级管路压力稳定 / Vacuum foreline pressure stabilization
  分类 Category : DL_Process
  码位 Code     : 16#06_0_99
  版本 Version  : 1.0.0
  溯源 Source   : ModPID 语义借鉴 · clean-room 实现，仅借分类/参数域/命名，未复制源码
  功能 Function : 1) 前级压力闭环 PI 调节（复用 FB_DL_PidController，阀位限幅抗饱和联动）；
                  2) 抽速前馈通道叠加（前馈指令非有限拒绝并保持末次有效）；
                  3) 压力越窗分级告警（带迟滞）。
  边界 Boundary : ① 压力无效冻结输出（跟踪回投保持末次阀位）；
                  ② 设定低于量程下限钳定并置码；
                  ③ 阀位饱和与 PI 抗饱和联动（限幅反算由实例承担）；
                  ④ 前馈通道指令非有限拒绝保持末次有效（FB_DL_SuperimposedMove 同范式）；
                  ⑤ 越窗分级带迟滞；
                  ⑥ 输出三行同向：阀位 → 饱和/冻结标志 → 越窗告警。
  依赖 Depends  : FB_DL_PidController × 1（PI 调节，每拍无条件调用）

  码表 Error codes（本件子码步进 16#30 · 本格 99 与既有 9X 子码段冲突，错位至 C9/D9 避让）:
    16#0002_06C9 故障级：组态非法（量程域倒置 / 行程域倒置 / 增益 <= 0）
    16#0002_06D9 故障级：相 ID 越界（枚举兜底路径）
    16#0002_06B9 信息级：压力无效输出冻结 / 设定低于量程钳定 / 前馈非有限已拒 / 越窗提示（不置 bError）
*)

TYPE E_DL_FpcPhase :
(
    eIdle   := 0,  // 空闲（阀位回下限）/ Idle, valve at low limit
    eRun    := 10, // PI 调节运行 / PI running
    eFrozen := 20, // 压力无效冻结 / Frozen by invalid pressure
    eFault  := 90  // 组态故障锁定 / Configuration fault locked
);
END_TYPE

FUNCTION_BLOCK FB_DL_ForelinePressureCtrl
VAR_INPUT
    bEnable       : BOOL;                           // 总使能，FALSE 阀位回下限 / Master enable
    bReset        : BOOL;                           // 复位，上升沿清组态故障 / Reset, clears fault
    fPressPa      : REAL;                           // 前级压力实测 [Pa] / Foreline pressure [Pa]
    fPressSpPa    : REAL := 10.0;                   // 压力设定 [Pa]，域 > 0 / Pressure setpoint [Pa]
    fRangeLoPa    : REAL := 1.0;                    // 量程下限 [Pa]，域 > 0（设定钳定域）/ Range low [Pa]
    fRangeHiPa    : REAL := 1000.0;                 // 量程上限 [Pa]，域 > 0 / Range high [Pa]
    fSpeedFfPct   : REAL;                           // 抽速前馈指令 [%] / Pumping-speed feedforward [%]
    fKp           : REAL := 2.0;                    // 比例增益 [1]，负值 = 反作用 / Proportional gain [1]
    tTi           : TIME := T#30S;                  // 积分时间 [s]，T#0S = 关闭 / Integral time, T#0S = off
    tTd           : TIME := T#0S;                   // 微分时间 [s]，T#0S = 关闭 / Derivative time, T#0S = off
    fValveMinPct  : REAL := 0.0;                    // 阀位行程域下限 [%] / Valve domain low [%]
    fValveMaxPct  : REAL := 100.0;                  // 阀位行程域上限 [%] / Valve domain high [%]
    fDevWarnPa    : REAL := 3.0;                    // 越窗提示门限 [Pa]，域 > 0 / Deviation warning limit [Pa]
    fHystPa       : REAL := 0.5;                    // 越窗迟滞 [Pa]，域 > 0 / Deviation hysteresis [Pa]
    fEps          : REAL := 1.0E-6;                 // 浮点判零容差 [1] / Floating zero tolerance
END_VAR
VAR_OUTPUT
    fValveOutPct  : REAL;                           // 调节阀位输出 [%]（PI + 前馈叠加）/ Valve output [%]
    fFfUsedPct    : REAL;                           // 本拍生效前馈 [%] / Feedforward used [%]
    bSaturated    : BOOL;                           // 阀位饱和标志 / Valve saturated flag
    bFrozen       : BOOL;                           // 压力无效冻结标志 / Frozen by invalid pressure
    bDevWarn      : BOOL;                           // 越窗提示标志（带迟滞）/ Deviation warning flag
    bError        : BOOL;                           // 故障标志，与故障级码配对 / Fault flag
    uErrorId      : UDINT;                          // 事件码，0 = 无事件 / Event code
    eStateOut     : E_DL_FpcPhase;                  // 状态机当前态，段尾单点映射 / Phase mapped at tail
END_VAR
VAR
    _eState       : E_DL_FpcPhase := E_DL_FpcPhase.eIdle;  // 内部状态 / Internal state
    fbPid         : FB_DL_PidController;            // PI 实例（无条件调用）/ PI instance
    rtrReset      : R_TRIG;                         // 复位沿 / Reset edge
    bCfgOk        : BOOL;                           // 组态合法标志 / Configuration valid
    bPressOk      : BOOL;                           // 压力本拍有效 / Pressure valid this scan
    fSpClampPa    : REAL;                           // 钳定后设定 [Pa] / Clamped setpoint [Pa]
    bSpClamped    : BOOL;                           // 设定钳定标志 / Setpoint clamped flag
    fFfHoldPct    : REAL;                           // 末次有效前馈 [%]（非有限保持）/ Last valid feedforward [%]
    bFfOk         : BOOL;                           // 前馈指令本拍有效 / Feedforward valid this scan
    bDevUp        : BOOL;                           // 越窗迟滞状态（持有）/ Deviation hysteresis state
    fValveHold    : REAL;                           // 末次有效阀位 [%]（冻结保持）/ Last valid valve [%]
    uFault        : UDINT;                          // 锁存故障码 / Latched fault code
    uInfo         : UDINT;                          // 信息级码 / Information code
END_VAR

(* === 段 0 · 实例刷新 === *)
rtrReset(CLK := bReset);                          // 每拍刷新复位沿

(* === 段 1 · 组态闸 === *)
bCfgOk := (fRangeHiPa > fRangeLoPa + fEps)        // 量程域不倒置
          AND (fValveMaxPct > fValveMinPct + fEps)// 行程域不倒置
          AND (ABS(fKp) > fEps)                   // 增益非零（负值 = 反作用合法）
          AND (fDevWarnPa > fHystPa)              // 越窗门限大于迟滞（带不相交）
          AND (fPressSpPa = fPressSpPa) AND (fKp = fKp);  // NaN 自反
IF NOT bCfgOk THEN
    uFault := 16#0002_06C9;                       // 故障级：组态非法
END_IF
IF rtrReset.Q AND bCfgOk THEN
    uFault := 16#0000;                            // 复位沿清锁存（解除路径可达）
    bDevUp := FALSE;                              // 越窗迟滞复位
END_IF
uInfo := 16#0000;                                 // 信息码每拍清零
bPressOk := (fPressPa = fPressPa) AND (fPressPa >= 0.0) AND (fPressPa < 1.0E30);   // 压力 NaN 自反 + 非负域闸

(* === 段 2 · 设定钳定与越窗迟滞判据（本拍重算）=== *)
fSpClampPa := fPressSpPa;                         // 设定先取组态值
bSpClamped := bPressOk AND (fSpClampPa < fRangeLoPa);   // 低于量程下限钳定标志
IF bSpClamped THEN
    fSpClampPa := fRangeLoPa;                     // 钳定量程下限
    uInfo := 16#0002_06B9;                        // 信息级：设定低于量程钳定
END_IF
bDevUp := bDevUp AND bPressOk;                    // 迟滞状态只在有效拍保持（无效拍判据挂起）
IF bPressOk THEN
    IF ABS(fPressPa - fSpClampPa) >= fDevWarnPa THEN
        bDevUp := TRUE;                           // 越窗置迟滞状态
    ELSIF ABS(fPressPa - fSpClampPa) < fDevWarnPa - fHystPa THEN
        bDevUp := FALSE;                          // 回差带内解除（路径可达）
    END_IF
END_IF
bDevWarn := bDevUp;                               // 越窗提示出口

(* === 段 3 · 前馈通道非有限拒绝（保持末次有效，SuperimposedMove 同范式）=== *)
bFfOk := (fSpeedFfPct = fSpeedFfPct) AND (ABS(fSpeedFfPct) < 1.0E30);   // 前馈 NaN 自反 + 幅值闸
IF bFfOk THEN
    fFfHoldPct := fSpeedFfPct;                    // 有效拍记账末次前馈
ELSE
    uInfo := 16#0002_06B9;                        // 信息级：前馈非有限已拒
END_IF
fFfUsedPct := fFfHoldPct;                         // 生效前馈（保持末次有效）

(* === 段 4 · PI 实例（每拍无条件调用，限幅反算抗饱和由实例承担）=== *)
fbPid(bEnable := bEnable AND bCfgOk AND bPressOk, // 压力无效/故障：PI 停调
      bManual := FALSE,                           // 自动调节
      fSetpoint := fSpClampPa,                    // 钳定后设定
      fActual := fPressPa,                        // 压力实测
      fKp := fKp,                                 // 比例增益
      tTi := tTi,                                 // 积分时间（0 = 关闭，合法语义）
      tTd := tTd,                                 // 微分时间（0 = 关闭）
      rOutMin := fValveMinPct - fFfUsedPct,       // 输出下限平移（前馈叠加域）
      rOutMax := fValveMaxPct - fFfUsedPct,       // 输出上限平移（前馈叠加域，限幅反算）
      tSampleTime := T#100MS,                     // 采样周期
      bTrack := (NOT bPressOk) OR (NOT bEnable),  // 无效/失能：跟踪回投保持阀位（无扰冻结）
      fTrackValue := fValveHold - fFfUsedPct,     // 跟踪值 = 末次阀位 − 前馈（叠加域口径）
      bReset := rtrReset.Q);                      // 复位沿透传
fValveOutPct := fbPid.fOut + fFfUsedPct;          // 阀位 = PI 输出 + 前馈叠加
IF fValveOutPct > fValveMaxPct THEN
    fValveOutPct := fValveMaxPct;                 // 钳到行程域上限
END_IF
IF fValveOutPct < fValveMinPct THEN
    fValveOutPct := fValveMinPct;                 // 钳到行程域下限
END_IF
bSaturated := fbPid.bLimitHigh OR fbPid.bLimitLow;   // 饱和标志（映射实例触限）
IF bSaturated AND bPressOk THEN
    uInfo := 16#0002_06B9;                        // 信息级：阀位饱和
END_IF

(* === 段 5 · 主状态机（ENUM + CASE，含 ELSE 兜底）=== *)
CASE _eState OF
E_DL_FpcPhase.eIdle :
    IF uFault <> 16#0000 THEN
        _eState := E_DL_FpcPhase.eFault;          // 故障优先
    ELSIF bEnable AND bCfgOk AND (NOT bPressOk) THEN
        _eState := E_DL_FpcPhase.eFrozen;         // 压力无效进冻结
    ELSIF bEnable AND bCfgOk AND bPressOk THEN
        _eState := E_DL_FpcPhase.eRun;            // 进运行相
    END_IF

E_DL_FpcPhase.eRun :
    IF (uFault <> 16#0000) OR (NOT bEnable) THEN
        _eState := E_DL_FpcPhase.eFault;          // 故障/失能转出
    ELSIF NOT bPressOk THEN
        uInfo := 16#0002_06B9;                    // 信息级：压力无效输出冻结
        _eState := E_DL_FpcPhase.eFrozen;         // 转冻结相（阀位保持末次值）
    ELSE
        fValveHold := fValveOutPct;               // 有效拍记账末次阀位（冻结保持源）
    END_IF

E_DL_FpcPhase.eFrozen :
    IF bPressOk AND bEnable AND (uFault = 16#0000) THEN
        _eState := E_DL_FpcPhase.eRun;            // 压力恢复回运行（解除路径可达，跟踪无扰）
    END_IF

E_DL_FpcPhase.eFault :
    IF uFault = 16#0000 THEN
        _eState := E_DL_FpcPhase.eIdle;           // 解锁回空闲
    END_IF

ELSE
    _eState := E_DL_FpcPhase.eFault;              // 非法状态拦截
    uFault := 16#0002_06D9;                       // 故障级：相 ID 越界
END_CASE
bFrozen := (_eState = E_DL_FpcPhase.eFrozen);     // 冻结标志段尾单点映射

(* === 段 6 · 输出映射 === *)
bError := (uFault <> 16#0000);                    // 故障标志仅由故障级码置位（R45 配对）
IF bError THEN
    uErrorId := uFault;                           // 故障级优先上报
ELSE
    uErrorId := uInfo;                            // 否则上报信息级码
END_IF
eStateOut := _eState;                             // 输出枚举段尾单点映射（N2 规则）
END_FUNCTION_BLOCK

(* ---- FB_DL_ForgeDieLubeSeq.st ---- *)
(*
  Name: FB_DL_ForgeDieLubeSeq
  Category: DL_Process
  Version: 1.0.0
  Round: R89 / 2026-11-25
  开源溯源：clean-room 自研（族 锻造加热退火，ST 开源生态实测 0 命中，无外部代码引入）
  功能：锻模润滑喷涂顺序：吹扫→喷涂→吹干→允许锻造，三段时长各自独立 TON。
  边界条件：① 三段时长为 TIME 入参，必须 > 0，否则组态非法（101）立即锁故障；
            ② 吹扫/喷涂/吹干各用独立 TON，PT 分别取 tBlowS / tSprayS / tDryS，禁跨相共用（R100 无同拍双窗）；
            ③ 气源不足（xAirOk = FALSE）在启动申请存在时即锁故障（102），并撤喷涂与锻造许可；
            ④ 故障解除唯一路径：故障相内 xStart 释放（R152），清锁存回 eIdle。
  状态机：eIdle / eBlow / eSpray / eDry / eReady / eFault（CASE 含 ELSE 兜底）。
*)
TYPE E_DL_DlsPhase :
(
    eIdle  := 0,        (* 待机：等启动沿 / Idle, waiting for start edge *)
    eBlow  := 10,       (* 吹扫相：压缩空气吹净型腔 / Blow phase, air purge *)
    eSpray := 20,       (* 喷涂相：润滑剂喷涂 / Spray phase, lubricant *)
    eDry    := 30,      (* 吹干相：吹干残留 / Dry phase, air dry *)
    eReady := 40,       (* 锻造许可相：允许锻造 / Forge permit phase *)
    eFault := 90        (* 故障相：锁存待释放 / Fault latched, awaiting release *)
);
END_TYPE

FUNCTION_BLOCK FB_DL_ForgeDieLubeSeq
VAR_INPUT
    xStart : BOOL;      (* 启动命令（上升沿起序） [-] Start command, rising edge *)
    tBlowS : TIME;      (* 吹扫时长 [ms] Blow duration [ms] *)
    tSprayS : TIME;     (* 喷涂时长 [ms] Spray duration [ms] *)
    tDryS : TIME;       (* 吹干时长 [ms] Dry duration [ms] *)
    xAirOk : BOOL;      (* 气源压力正常 [-] Air supply healthy *)
END_VAR
VAR_OUTPUT
    eState : E_DL_DlsPhase;  (* 当前相 [-] Present phase *)
    xSprayValve : BOOL;      (* 喷涂阀指令（仅喷涂相） [-] Spray valve command *)
    xAllowForge : BOOL;      (* 允许锻造 [-] Forge permitted *)
    xFault : BOOL;           (* 故障锁存标志 [-] Fault latched *)
END_VAR
VAR
    _ePhase : E_DL_DlsPhase := E_DL_DlsPhase.eIdle;  (* 内部相（CASE 唯一写入目标） [-] Internal phase *)
    _bFaultLatch : BOOL := FALSE;   (* 故障锁存位 [-] Fault latch *)
    _bReqFault : BOOL := FALSE;     (* 单拍故障请求（段 1 预清） [-] Fault request *)
    tonBlow : TON;                  (* 吹扫计时（段 0 无条件调用） / Blow timer *)
    tonSpray : TON;                 (* 喷涂计时（段 0 无条件调用） / Spray timer *)
    tonDry : TON;                   (* 吹干计时（段 0 无条件调用） / Dry timer *)
    rtStart : R_TRIG;               (* 启动沿（段 0 无条件调用） / Start edge *)
END_VAR
(* —— 段 0：沿与三 TON 无条件周期刷新（R7），IN 仅由相位派生 —— *)
rtStart(CLK := xStart);                                             (* 启动沿 / Start edge *)
tonBlow(IN := (_ePhase = E_DL_DlsPhase.eBlow), PT := tBlowS);       (* 吹扫计时 / Blow timer *)
tonSpray(IN := (_ePhase = E_DL_DlsPhase.eSpray), PT := tSprayS);    (* 喷涂计时 / Spray timer *)
tonDry(IN := (_ePhase = E_DL_DlsPhase.eDry), PT := tDryS);          (* 吹干计时 / Dry timer *)
(* —— 段 1：单拍量预清 + 组态/气源故障请求（本件无码出口，成因由相位 + xFault 表达） —— *)
_bReqFault := FALSE;
IF (tBlowS <= T#0S) OR (tSprayS <= T#0S) OR (tDryS <= T#0S) THEN
    _bReqFault := TRUE;                         (* 组态非法：时长为零 / Configuration bad, zero duration *)
ELSIF xStart AND (NOT xAirOk) THEN
    _bReqFault := TRUE;                         (* 气源不足 / Air supply low *)
END_IF
(* —— 段 2：故障锁存解除（唯一路径 = 故障相内 xStart 释放，R152） —— *)
IF _bFaultLatch AND (NOT xStart) THEN
    _bFaultLatch := FALSE;                      (* 清锁存 / Clear latch *)
    _ePhase := E_DL_DlsPhase.eIdle;             (* 迁回待机 / Back to idle *)
END_IF
(* —— 段 3：主状态机（ENUM + CASE，ELSE 兜底） —— *)
CASE _ePhase OF
E_DL_DlsPhase.eIdle:
    IF rtStart.Q AND (NOT _bFaultLatch) AND xAirOk THEN
        _ePhase := E_DL_DlsPhase.eBlow;         (* 起序 → 吹扫 / Start, blow *)
    END_IF
E_DL_DlsPhase.eBlow:
    IF tonBlow.Q THEN
        _ePhase := E_DL_DlsPhase.eSpray;        (* 吹扫到时 → 喷涂 / Blow done, spray *)
    END_IF
E_DL_DlsPhase.eSpray:
    IF tonSpray.Q THEN
        _ePhase := E_DL_DlsPhase.eDry;          (* 喷涂到时 → 吹干 / Spray done, dry *)
    END_IF
E_DL_DlsPhase.eDry:
    IF tonDry.Q THEN
        _ePhase := E_DL_DlsPhase.eReady;        (* 吹干到时 → 许可锻造 / Dry done, permit *)
    END_IF
E_DL_DlsPhase.eReady:
    IF NOT xStart THEN
        _ePhase := E_DL_DlsPhase.eIdle;         (* 启动释放 → 待机（撤许可） / Start released *)
    END_IF
E_DL_DlsPhase.eFault:
    _bReqFault := FALSE;                        (* 故障相驻留：锁存已置，不再新发请求 *)
ELSE
    _bReqFault := TRUE;                         (* 非法相兜底 / Illegal phase fallback *)
END_CASE
(* —— 段 4：故障请求统一落地（唯一锁存点 + 同步迁相，R187/R252） —— *)
IF _bReqFault AND (NOT _bFaultLatch) THEN
    _bFaultLatch := TRUE;                       (* 锁存 / Latch *)
    _ePhase := E_DL_DlsPhase.eFault;            (* 同步迁相 / Migrate to fault *)
END_IF
(* —— 段 5：统一出口（各出口单点赋值） —— *)
eState := _ePhase;
xSprayValve := (_ePhase = E_DL_DlsPhase.eSpray) AND (NOT _bFaultLatch);
xAllowForge := (_ePhase = E_DL_DlsPhase.eReady) AND (NOT _bFaultLatch) AND xAirOk;
xFault := _bFaultLatch;
END_FUNCTION_BLOCK

(* ---- FB_DL_FormationChannelMgr.st ---- *)
//==============================================================================
// 功能块：FB_DL_FormationChannelMgr ｜ 中文名称：化成/分容柜通道调度
// 所属子库：DL_Process ｜ 版本：v1.0.0 ｜ 兼容：CODESYS V3.5+ / TwinCAT 3 / 汇川 InoProShop
// 功能描述：化成/分容柜多通道调度：空闲通道分配（跳过隔离与故障通道）→ 批次启动命令 →
//           异常通道隔离锁存 → 批次完成/中止 → 台账计数（完成数/故障数）。
//           本件只做「调度层」，绝不内联充放电工步机（工步归序号 15 的 BatteryTestCycler）：
//           两者以布尔快照（abChBusy / abChFault / abChDone）与指令握手位
//           （abChCmdStart）交互，本件不产生任何电流/电压设定，也不判任何工艺终止条件。
//           无空闲通道属产线常态，挂起等待并给信息码，绝不升格为故障。
// 开源溯源 (Origin)：道莅原创实现（参考 公开工程惯例 分类与参数域）
// 单位表：通道数[路] / 通道号[号] / 计数[路] / 布尔快照[—]
// 错误码表：16#0005_040E 信息级（无空闲通道，分配挂起，不置 bError）/
//           16#0005_040F 信息级（异常通道已隔离并记账，锁存至 bReset，不置 bError）/
//           16#0005_0357 故障级（通道数非法/数组域越界，置 bError）/ 16#0005_0358
//           故障级（重复分配：上一分配尚未启动又发新请求，防双工步叠加烧电芯，置 bError）/
//           16#0005_0359 故障级兜底（状态机落 ELSE 非法状态，置 bError）。码位 16#0005 段。
// 状态机：E_DL_FormationChState（eIdle=0 待机 / eStandby=10 可分配待命 / eBatchRun=20
//           批次运行 / eBatchDone=30 批次完成 / eFault=99 故障兜底），CASE 含 ELSE 兜底，
//           ELSE 置 0359 且撤全通道启动指令、许可撤。
// 边界行为：① 无空闲通道 → bAllocOk := FALSE + 信息 040E，挂起等待不置故障（产线常态）；
//           ② 故障通道 → 隔离锁存 abChBlocked + 信息 040F（锁存至 bReset，防止自动复用
//           坏通道）；③ nChannelCount 域 1~16，越界 → 故障 0357；④ 上一分配未启动又发
//           新分配请求 → 故障 0358（防同一通道双工步叠加）；⑤ bBatchAbort → 撤全通道
//           启动指令 + bBatchAborted（中止优先于完成）；⑥ 失能 → 撤指令 + bValid := FALSE
//           （R72）；⑦ 数组一律按 nChannelCount 上界遍历（域已闸），不做越界下标访问。
// 修订历史：v1.0.0 2026-11-17 首版（R25 派单 · §4.19，与 §4.15 件布尔握手分层）
//==============================================================================
(*------------------------------------------------------------------------------
 * 枚举: E_DL_FormationChState（归属 DL_Process，与 FB_DL_FormationChannelMgr 同文件）
 *----------------------------------------------------------------------------*)
TYPE E_DL_FormationChState :
(
    eIdle      := 0,   // 待机：失能，全通道启动指令撤 / Idle, all channel start commands dropped
    eStandby   := 10,  // 待命：可接受分配请求 / Standby, allocation requests accepted
    eBatchRun  := 20,  // 批次运行：已启动通道在跑 / Batch running
    eBatchDone := 30,  // 批次完成：全部已启动通道报完成 / Batch completed
    eFault     := 99   // 故障兜底：通道数非法/重复分配/非法状态 / Fault fallback
);
END_TYPE

(*==============================================================================
 * 功能块: FB_DL_FormationChannelMgr
 * 调用约定: 每个扫描周期无条件调用一次；通道快照由柜体通信层刷新。
 *============================================================================*)
FUNCTION_BLOCK FB_DL_FormationChannelMgr
VAR_INPUT
    abChBusy         : ARRAY[0..15] OF BOOL;       // 通道忙快照（柜体层刷新）/ Channel busy snapshot
    abChFault        : ARRAY[0..15] OF BOOL;       // 通道故障快照 / Channel fault snapshot
    abChDone         : ARRAY[0..15] OF BOOL;       // 通道完成快照 / Channel done snapshot
    nChannelCount    : INT := 16;                  // 有效通道数 [路]，合法域 1~16 / Usable channel count, domain 1..16
    bAllocReq        : BOOL;                       // 分配请求（取上升沿）/ Allocation request, rising edge
    bBatchStart      : BOOL;                       // 批次启动（取上升沿）/ Batch start, rising edge
    bBatchAbort      : BOOL;                       // 批次中止（取上升沿，优先于完成）/ Batch abort, rising edge, outranks completion
    bEnable          : BOOL;                       // 总使能 / Master enable
    bReset           : BOOL;                       // 复位，上升沿清隔离锁存与台账 / Reset, rising edge clears the isolation latches and the ledger
END_VAR
VAR_OUTPUT
    nAllocatedCh     : INT;                        // 已分配通道号 [号]，-1 = 未分配 / Allocated channel, -1 = none
    bAllocOk         : BOOL;                       // 分配成功（单拍脉冲）/ Allocation succeeded, single-scan pulse
    abChBlocked      : ARRAY[0..15] OF BOOL;       // 通道隔离掩码（锁存至 bReset）/ Channel isolation mask, latched
    abChCmdStart     : ARRAY[0..15] OF BOOL;       // 通道启动指令 / Channel start command
    nDoneCount       : INT;                        // 完成通道数 [路] / Completed channels
    nFaultCount      : INT;                        // 故障通道数 [路] / Faulted channels
    bBatchDone       : BOOL;                       // 批次完成 / Batch completed
    bBatchAborted    : BOOL;                       // 批次已中止 / Batch aborted
    eErr             : UDINT;                      // 错误码，0 = 无错，码位 16#0005_040E 起信息级、16#0005_0357 起故障级（分带见错误码表） / Error code, 0 = no error, band info/fault per the code table
    bError           : BOOL;                       // 故障级标志，仅故障级错误置位 / Fault-class flag, set only on fault-level codes
    bValid           : BOOL;                       // 调度输出可用标志，失能/故障闸显式 FALSE / Schedule usable flag, explicit FALSE on disable/fault gates
    eState           : E_DL_FormationChState;      // 主状态机当前状态 / Current state of the main state machine
END_VAR
VAR
    fbReset          : R_TRIG;                     // 复位上升沿检测实例 / Reset rising edge detector
    fbAlloc          : R_TRIG;                     // 分配请求上升沿检测实例 / Allocation request rising edge detector
    fbStart          : R_TRIG;                     // 批次启动上升沿检测实例 / Batch start rising edge detector
    fbAbort          : R_TRIG;                     // 批次中止上升沿检测实例 / Batch abort rising edge detector
    abCmdInt         : ARRAY[0..15] OF BOOL;       // 启动指令内部副本 / Internal command copy
    nLoop            : INT;                        // 遍历索引 [—] / Loop index
    nFreeCh          : INT;                        // 候选空闲通道号 [号] / Candidate free channel
    bAllocPending    : BOOL;                       // 已分配但尚未启动（重复分配判据）/ Allocated but not started, the duplicate-allocation predicate
    bIsoNew          : BOOL;                       // 本拍新隔离通道标志 / A channel was newly isolated this scan
    bAnyCmd          : BOOL;                       // 存在启动指令 / Any start command active
    bAllDone         : BOOL;                       // 已启动通道全部报完成 / Every started channel reports done
    bNonFree         : BOOL;                       // 本拍无空闲通道 / No free channel this scan
    bFirstScan       : BOOL := TRUE;               // 上电首拍标志 / First-scan flag
END_VAR
VAR CONSTANT
    DL_FCM_CODE_INFO_1 : UDINT := 16#0005_040E;    // 信息级槽 1（无空闲通道，分配挂起） / info slot 1
    DL_FCM_CODE_INFO_2 : UDINT := 16#0005_040F;    // 信息级槽 2（异常通道已隔离并记账） / info slot 2
    DL_FCM_CODE_FLT_1  : UDINT := 16#0005_0357;    // 故障级槽 1（通道数非法/数组域越界） / fault slot 1
    DL_FCM_CODE_FLT_2  : UDINT := 16#0005_0358;    // 故障级槽 2（重复分配） / fault slot 2
    DL_FCM_CODE_FLT_3  : UDINT := 16#0005_0359;    // 故障级槽 3（非法状态兜底） / fault slot 3
    DL_FCM_CH_MAX      : INT := 16;                // 通道上限 [路]，必须等于数组维度 / Channel ceiling, must match the arrays
    DL_FCM_CH_MIN      : INT := 1;                 // 通道下限 [路] / Channel floor
    DL_FCM_IDX_NONE    : INT := -1;                // 无效通道号哨兵 [号] / Invalid channel sentinel
END_VAR

(*------------------------------------------------------------------------------
 * 段 1｜无条件刷新区（红线 5）：四条沿检测在任意分支之外周期调用
 *----------------------------------------------------------------------------*)
bAllocOk := FALSE;                                 // 分配成功为单拍脉冲，逐拍先清 / single-scan pulse cleared first
fbReset(CLK := bReset);                            // 复位沿检测无条件刷新 / reset edge refreshed unconditionally
fbAlloc(CLK := bAllocReq);                         // 分配请求沿检测无条件刷新 / allocation edge refreshed unconditionally
fbStart(CLK := bBatchStart);                       // 批次启动沿检测无条件刷新 / start edge refreshed unconditionally
fbAbort(CLK := bBatchAbort);                       // 批次中止沿检测无条件刷新 / abort edge refreshed unconditionally

(*------------------------------------------------------------------------------
 * 段 2｜复位沿处理（改写置于沿后，防吞沿 R39）：清隔离锁存与台账
 *----------------------------------------------------------------------------*)
IF fbReset.Q THEN
    eState := E_DL_FormationChState.eIdle;
    eErr   := 16#0000_0000;                        // 复位清码 / reset clears the code
    bError := FALSE;                               // 复位清故障 / reset clears the fault
    bBatchDone := FALSE;                           // 批次完成标志清 / batch-done flag cleared
    bBatchAborted := FALSE;                        // 中止标志清 / aborted flag cleared
    bAllocPending := FALSE;                        // 待启动分配清 / pending allocation cleared
    nDoneCount := 0;                               // 完成计数清 / done count cleared
    nFaultCount := 0;                              // 故障计数清 / fault count cleared
    nAllocatedCh := DL_FCM_IDX_NONE;               // 分配通道清 / allocated channel cleared
    FOR nLoop := 0 TO DL_FCM_CH_MAX - 1 DO
        abChBlocked[nLoop] := FALSE;               // 隔离锁存清除 / isolation latch cleared
        abCmdInt[nLoop] := FALSE;                  // 启动指令内部副本清 / internal command cleared
        abChCmdStart[nLoop] := FALSE;              // 启动指令出口清 / command outlet cleared
    END_FOR
    bFirstScan := TRUE;                            // 重新首拍化 / re-initialize first scan
END_IF

(*------------------------------------------------------------------------------
 * 段 3｜通道数域闸（先闸后遍历：后续所有循环都以 nChannelCount 为上界）
 *----------------------------------------------------------------------------*)
IF (nChannelCount < DL_FCM_CH_MIN) OR (nChannelCount > DL_FCM_CH_MAX) THEN
    eState := E_DL_FormationChState.eFault;        // 进故障相 / enter fault state
    eErr   := DL_FCM_CODE_FLT_1;                   // 故障级：通道数非法/数组域越界 / fault: channel count out of range
    bError := TRUE;                                // 故障级必置 bError（R45 配对）/ fault-class pairs with bError
    bValid := FALSE;                               // 调度不可用 / schedule unusable
    bAllocOk := FALSE;                             // 分配不成立 / allocation void
    nAllocatedCh := DL_FCM_IDX_NONE;               // 通道号清 / channel cleared
    FOR nLoop := 0 TO DL_FCM_CH_MAX - 1 DO
        abChCmdStart[nLoop] := FALSE;              // 全撤启动指令安全侧 / every command dropped
    END_FOR
    RETURN;
END_IF

(*------------------------------------------------------------------------------
 * 段 4｜通道隔离记账（锁存至 bReset）：故障通道一经发现立即隔离，
 *       并计入故障台账；隔离是「不再自动复用坏通道」的唯一手段
 *----------------------------------------------------------------------------*)
bIsoNew := FALSE;                                  // 本拍隔离标志初值 / isolation seed
nFaultCount := 0;                                  // 故障计数重数 / fault count recounted
FOR nLoop := 0 TO nChannelCount - 1 DO
    IF abChFault[nLoop] THEN
        nFaultCount := nFaultCount + 1;            // 故障通道计数 [路] / faulted channel counted
        IF NOT abChBlocked[nLoop] THEN
            abChBlocked[nLoop] := TRUE;            // 隔离锁存（首次）/ isolation latched on first detection
            bIsoNew := TRUE;                       // 本拍有新隔离 / newly isolated this scan
        END_IF
    END_IF
END_FOR

(*------------------------------------------------------------------------------
 * 段 5｜重复分配闸：上一分配已占通道但尚未启动批次，又来新的分配请求 → 0358
 *       （同一通道被两次工步叠加会烧电芯，属安全级）
 *----------------------------------------------------------------------------*)
IF fbAlloc.Q AND bAllocPending THEN
    eState := E_DL_FormationChState.eFault;        // 进故障相 / enter fault state
    eErr   := DL_FCM_CODE_FLT_2;                   // 故障级：重复分配 / fault: duplicate allocation
    bError := TRUE;                                // 故障级必置 bError（R45 配对）/ fault-class pairs with bError
    bValid := FALSE;                               // 调度不可用 / schedule unusable
    bAllocOk := FALSE;                             // 分配不成立 / allocation void
    FOR nLoop := 0 TO nChannelCount - 1 DO
        abChCmdStart[nLoop] := FALSE;              // 全撤启动指令安全侧 / every command dropped
    END_FOR
    RETURN;
END_IF

(*------------------------------------------------------------------------------
 * 段 6｜分配：首个「未忙、未隔离、无故障」通道；无空闲 → 040E 挂起（不置故障）
 *----------------------------------------------------------------------------*)
nFreeCh := DL_FCM_IDX_NONE;                        // 候选通道初值 / candidate seed
FOR nLoop := 0 TO nChannelCount - 1 DO
    IF (NOT abChBlocked[nLoop]) AND (NOT abChFault[nLoop]) AND (NOT abChBusy[nLoop])
       AND (nFreeCh = DL_FCM_IDX_NONE) THEN
        nFreeCh := nLoop;                          // 取首个「未忙、未隔离、无故障」通道 [号] / first free channel wins
    END_IF
END_FOR
bNonFree := (nFreeCh = DL_FCM_IDX_NONE);           // 无空闲通道判据 / no-free-channel predicate
IF fbAlloc.Q AND (NOT bAllocPending) THEN
    IF bNonFree THEN
        bAllocOk := FALSE;                         // 分配不成立（挂起）/ allocation suspended
        nAllocatedCh := DL_FCM_IDX_NONE;           // 通道号保持无效 / channel stays invalid
        eErr := DL_FCM_CODE_INFO_1;                // 信息级：无空闲通道，分配挂起（产线常态，不置故障）/ info: no free channel, suspended
        bError := FALSE;                           // 信息级不置 bError（R45/R101）/ info never raises bError
    ELSE
        nAllocatedCh := nFreeCh;                   // 落定分配通道 [号] / the allocation settles
        bAllocOk := TRUE;                          // 分配成功单拍脉冲 / single-scan success pulse
        bAllocPending := TRUE;                     // 待启动（重复分配判据置位）/ pending, the duplicate predicate raises
        bBatchAborted := FALSE;                    // 新分配开启新批次：中止标志撤 / a new allocation clears the abort flag
        bBatchDone := FALSE;                       // 新分配开启新批次：完成标志撤 / a new allocation clears the done flag
        eErr := 16#0000_0000;                      // 分配成功不占码位 / no code on success
        bError := FALSE;                           // 无故障 / no fault
    END_IF
END_IF

(*------------------------------------------------------------------------------
 * 段 7｜批次启动/中止握手：启动只作用于已分配通道；中止撤全部通道指令，
 *       且中止优先于完成判定（安全侧）
 *----------------------------------------------------------------------------*)
IF fbStart.Q AND bAllocPending AND (nAllocatedCh >= 0) AND (nAllocatedCh < nChannelCount) THEN
    abCmdInt[nAllocatedCh] := TRUE;                // 启动已分配通道 / start the allocated channel
    bAllocPending := FALSE;                        // 该分配已启动，解除待启动 / allocation consumed
    eState := E_DL_FormationChState.eBatchRun;     // 进批次运行相 / enter the batch-run state
END_IF
IF fbAbort.Q THEN
    FOR nLoop := 0 TO nChannelCount - 1 DO
        abCmdInt[nLoop] := FALSE;                  // 中止：撤全通道启动指令 / abort drops every command
    END_FOR
    bAllocPending := FALSE;                        // 待启动分配作废 / pending allocation voided
    bBatchAborted := TRUE;                         // 中止标志置位（优先于完成）/ aborted outranks done
    bBatchDone := FALSE;                           // 完成标志不得冒充 / done must not pose
    eState := E_DL_FormationChState.eStandby;      // 回待命 / back to standby
END_IF

(*------------------------------------------------------------------------------
 * 段 8｜完成判定：曾有指令且已启动通道全部报完成 → 批次完成（bBatchAborted 时不成立）
 *----------------------------------------------------------------------------*)
bAnyCmd := FALSE;                                  // 指令存在标志初值 / command-presence seed
bAllDone := TRUE;                                  // 全部完成判据初值 / all-done seed
FOR nLoop := 0 TO nChannelCount - 1 DO
    IF abCmdInt[nLoop] THEN
        bAnyCmd := TRUE;                           // 存在启动指令 / a command exists
        IF NOT abChDone[nLoop] THEN
            bAllDone := FALSE;                     // 有通道未完成 / a channel is not done
        END_IF
    END_IF
END_FOR
IF bAnyCmd AND bAllDone AND (NOT bBatchAborted) THEN
    bBatchDone := TRUE;                            // 批次完成 / batch completed
    eState := E_DL_FormationChState.eBatchDone;    // 进完成相 / enter the done state
    FOR nLoop := 0 TO nChannelCount - 1 DO
        abCmdInt[nLoop] := FALSE;                  // 完成即撤指令（工步机自会收尾）/ commands dropped on completion
    END_FOR
END_IF

(*------------------------------------------------------------------------------
 * 段 9｜台账计数：完成/故障通道数按 nChannelCount 上界遍历统计（域已闸）
 *----------------------------------------------------------------------------*)
nDoneCount := 0;                                   // 完成计数重数 / done count recounted
FOR nLoop := 0 TO nChannelCount - 1 DO
    IF abChDone[nLoop] THEN
        nDoneCount := nDoneCount + 1;              // 完成通道计数 [路] / completed channel counted
    END_IF
END_FOR

(*------------------------------------------------------------------------------
 * 段 10｜状态机：CASE 含 ELSE 兜底（非法状态 → 0359 + 全撤指令 + 许可撤）
 *----------------------------------------------------------------------------*)
CASE eState OF

    E_DL_FormationChState.eIdle:
        bValid := FALSE;                           // 失能闸显式不可用（R72）/ explicit FALSE on the disable gate
        bBatchDone := FALSE;                       // 完成标志撤 / done flag withdrawn
        bBatchAborted := FALSE;                    // 中止标志撤 / aborted flag withdrawn
        nAllocatedCh := DL_FCM_IDX_NONE;           // 分配通道清 / allocated channel cleared
        bAllocPending := FALSE;                    // 待启动分配清 / pending cleared
        eErr := 16#0000_0000;                      // 待机无错 / no error in idle
        bError := FALSE;                           // 待机无故障 / no fault in idle
        FOR nLoop := 0 TO DL_FCM_CH_MAX - 1 DO
            abCmdInt[nLoop] := FALSE;              // 待机撤指令 / commands dropped in idle
        END_FOR
        IF bEnable THEN
            eState := E_DL_FormationChState.eStandby;   // 使能进待命 / enable enters standby
            bFirstScan := FALSE;                   // 首拍标志清除 / first-scan flag cleared
        END_IF

    E_DL_FormationChState.eStandby:
        bValid := TRUE;                            // 调度可用 / schedule usable
        bError := FALSE;                           // 待命无故障 / no fault in standby
        IF bIsoNew THEN
            eErr := DL_FCM_CODE_INFO_2;            // 信息级：异常通道已隔离并记账 / info: channel isolated and booked
        ELSIF bNonFree AND fbAlloc.Q THEN
            eErr := DL_FCM_CODE_INFO_1;            // 信息级：无空闲通道，分配挂起 / info: no free channel, suspended
        ELSIF eErr <> DL_FCM_CODE_INFO_1 THEN
            eErr := 16#0000_0000;                  // 其余情况清码（挂起提示保持一拍）/ otherwise clear, keeping the hint for one scan
        END_IF
        IF NOT bEnable THEN
            eState := E_DL_FormationChState.eIdle; // 失能回待机 / disable returns to idle
            bValid := FALSE;                       // 失能闸显式不可用 / explicit FALSE on the disable gate
        END_IF

    E_DL_FormationChState.eBatchRun:
        bValid := TRUE;                            // 调度可用 / schedule usable
        bError := FALSE;                           // 运行相无故障 / no fault while running
        eErr := 16#0000_0000;                      // 运行相先清码 / clear the code first
        IF bIsoNew THEN
            eErr := DL_FCM_CODE_INFO_2;            // 信息级：异常通道已隔离 / info: channel isolated
        END_IF
        IF NOT bEnable THEN
            eState := E_DL_FormationChState.eIdle; // 失能回待机（退出条件一）/ disable, first exit
            bValid := FALSE;                       // 失能闸显式不可用 / explicit FALSE on the disable gate
            FOR nLoop := 0 TO nChannelCount - 1 DO
                abCmdInt[nLoop] := FALSE;          // 失能撤全部指令 / every command dropped
            END_FOR
        ELSIF NOT bAnyCmd THEN
            eState := E_DL_FormationChState.eStandby;   // 无指令回待命（退出条件二）/ no command left, second exit
        END_IF

    E_DL_FormationChState.eBatchDone:
        bValid := TRUE;                            // 完成台账可用 / the completed ledger is usable
        bBatchDone := TRUE;                        // 完成标志保持到下次分配 / done held until the next allocation
        bError := FALSE;                           // 完成相无故障 / no fault when done
        eErr := 16#0000_0000;                      // 完成无错 / no error when done
        IF NOT bEnable THEN
            eState := E_DL_FormationChState.eIdle; // 失能回待机（退出条件一）/ disable, first exit
            bValid := FALSE;                       // 失能闸显式不可用 / explicit FALSE on the disable gate
            bBatchDone := FALSE;                   // 完成标志撤 / done flag withdrawn
        ELSIF fbAlloc.Q THEN
            bBatchDone := FALSE;                   // 新分配即结束上一批（退出条件二）/ a new allocation closes the batch
            eState := E_DL_FormationChState.eStandby;   // 回待命 / back to standby
        END_IF

    E_DL_FormationChState.eFault:
        bValid := FALSE;                           // 故障闸显式不可用（R72）/ explicit FALSE on the fault gate
        bError := TRUE;                            // 故障级必置 bError（R45 配对）/ fault-class pairs with bError
        bAllocOk := FALSE;                         // 分配不成立 / allocation void
        bAllocPending := FALSE;                    // 待启动分配作废 / pending allocation voided
        FOR nLoop := 0 TO DL_FCM_CH_MAX - 1 DO
            abCmdInt[nLoop] := FALSE;              // 故障撤全通道指令（安全值而非上次值）/ every command dropped
        END_FOR
        IF eErr = 16#0000_0000 THEN
            eErr := DL_FCM_CODE_FLT_3;             // 入口无码时按非法状态兜底（R45：bError 必须有对应码）/ illegal-state fallback
        END_IF
        IF bEnable AND (nChannelCount >= DL_FCM_CH_MIN) AND (nChannelCount <= DL_FCM_CH_MAX) THEN
            eState := E_DL_FormationChState.eIdle; // 通道数合法且使能才回待机（退出条件 ≥2）/ recover only when the count is sane
        END_IF

    ELSE
        eState := E_DL_FormationChState.eFault;    // 非法状态兜底 / illegal-state fallback
        eErr := DL_FCM_CODE_FLT_3;                 // 故障级兜底：非法状态 / fault fallback: illegal state
        bError := TRUE;                            // 故障级必置 bError（R45 配对）/ fault-class pairs with bError
        bValid := FALSE;                           // 调度不可用 / schedule unusable
        bAllocOk := FALSE;                         // 分配不成立 / allocation void
        FOR nLoop := 0 TO DL_FCM_CH_MAX - 1 DO
            abCmdInt[nLoop] := FALSE;              // 全撤启动指令安全侧 / every command dropped
        END_FOR

END_CASE

(*------------------------------------------------------------------------------
 * 段 11｜出口装配：内部副本落到输出数组；失能/故障一律全撤（安全值而非上次值）
 *----------------------------------------------------------------------------*)
FOR nLoop := 0 TO DL_FCM_CH_MAX - 1 DO
    IF nLoop < nChannelCount AND bEnable AND bValid THEN
        abChCmdStart[nLoop] := abCmdInt[nLoop];    // 正常调度：透传内部副本 / pass the internal copy through
    ELSE
        abChCmdStart[nLoop] := FALSE;              // 失能/故障/域外：全撤安全侧 / drop everything, safe side
    END_IF
END_FOR
END_FUNCTION_BLOCK

(* ---- FB_DL_FormationChannelQueue.st ---- *)
(*==============================================================================
 * 组件名称 (Component)  : FB_DL_FormationChannelQueue
 * 所属子库 (Sublibrary) : DL_Process
 * 当前版本 (Version)    : 1.0.0
 * 兼容性 (Platform)     : CODESYS 3.5+ / TwinCAT 3 / 汇川 InoProShop / 施耐德 Machine Expert
 *                         仅依赖 Standard.library（R_TRIG / ABS），零厂商私有库
 * 功能描述 (Function)   : 化成柜通道排队与优先级抢占调度。申请（通道号+
 *                         优先级 0 高..3 低）入队；调度相取队列中最高优先级
 *                         （数值最小，同级先入先出）派发；运行中更高级申请到
 *                         来即抢占（当前通道回队头，bPreempt 单拍）；被派通道
 *                         bChanFault 电平即故障摘除（不回队，bEvict 单拍）；
 *                         bChanDone 沿正常收口计数。与 MotionCmdQueue/FifoBuffer
 *                         （通用队列）分工：本件是资源排队 + 优先级抢占 + 故障
 *                         摘除的调度语义。
 * 来源标签 (Origin)     : ROADMAP §16.1 R11 池（L694），自研 clean-room
 * 边界语义 (Boundary)   : ① 队满申请沿：bQueueFull 指示该拍拒收（申请丢弃，
 *                         头注释明示不缓存）；
 *                         ② 摘除/收口/抢占后的队列搬移用单向前移复制，游标
 *                         0..8 结构性有界；
 *                         ③ 优先级域闸 0..3 / 通道号域闸 1..99 越域 → 组态故障；
 *                         ④ 抢占只回队不重派，防同拍振荡。
 * 输出语义 (Fallback)   : 【R191】bEnable = FALSE → 派发保持（运行通道不中断，
 *                         由调用方决定停机）；eFault 相 → 派发撤销 + bError = TRUE。
 * 码位     (Codes)      : 按 R297 范式零 16# 码位硬编码；错误出口 BOOL+ENUM(eCause)。
 * 红线自检 (Redline)    : 7 项红线已自检：R1 零全局 ✓｜R2 零物理地址 ✓｜R3 纯 IEC ✓
 *                         R4 越界（游标有界）/组态闸 ✓｜R5 双语同行注释 ✓
 *                         R6 CASE 带 ELSE 兜底迁 eFault ✓｜R7 R_TRIG 段 0 无条件刷新 ✓
 * 验收向量 (Acceptance) : V1 队空申请（5,1）→ 立即派发 nDispatch=5；
 *                         V2 运行中申请（7,0）→ bPreempt 单拍，5 回队头，
 *                         7 抢占派发；
 *                         V3 运行通道故障电平 → bEvict 单拍不回队，自动派
 *                         队内次高优先级。
 * 修订历史 (Revision)   : 2026-11-20  v1.0.0  R51 首版（批 1 · 序号 3）
 *==============================================================================*)
TYPE E_DL_FcqState :
(
    eIdle  := 0,                             (* 待使能 / Idle *)
    eDispatch := 10,                         (* 有通道运行（队列可继续接纳） / Dispatching *)
    eFault := 90                             (* 故障锁存相 / Fault latched phase *)
);
END_TYPE

TYPE E_DL_FcqCause :
(
    eNone       := 0,                        (* 无故障成因 / No cause *)
    eCfgIllegal := 1,                        (* 组态非法：优先级/通道号越域 / Illegal config *)
    ePhaseBad   := 2                         (* 非法相位兜底 / Illegal phase fallback *)
);
END_TYPE

FUNCTION_BLOCK FB_DL_FormationChannelQueue
VAR_INPUT
    bReq       : BOOL := FALSE;              (* 申请电平（上升沿入队）[-] / Request level, edge enqueues *)
    nChanId    : INT := 0;                   (* 申请通道号，域 1..99 [-] / Channel id *)
    nPrio      : INT := 3;                   (* 申请优先级 0 高..3 低，域 0..3 [-] / Priority *)
    bChanDone  : BOOL := FALSE;              (* 运行通道完成沿 [-] / Dispatched channel done edge *)
    bChanFault : BOOL := FALSE;              (* 运行通道故障电平（摘除不回队）[-] / Dispatched channel fault *)
    bEnable    : BOOL := TRUE;               (* 使能 [-] / Enable *)
    bReset     : BOOL := FALSE;              (* 复位命令，上升沿清全部 [-] / Reset command *)
END_VAR
VAR_OUTPUT
    nDispatchId : INT;                       (* 派发通道号（0 = 无派发）[-] / Dispatched channel id *)
    bDispatchValid : BOOL;                   (* 派发有效指示 [-] / Dispatch valid *)
    nQueueDepth : INT;                       (* 当前队列深度 [条] / Queue depth *)
    bQueueFull  : BOOL;                      (* 队满指示（该拍申请拒收）[-] / Queue full *)
    bPreempt    : BOOL;                      (* 抢占单拍位 [-] / Preempt pulse *)
    bEvict      : BOOL;                      (* 故障摘除单拍位 [-] / Evict pulse *)
    nDoneCnt    : UDINT;                     (* 正常收口累计 [次] / Done count *)
    eState      : E_DL_FcqState;             (* 状态出口 / State outlet *)
    eCause      : E_DL_FcqCause;             (* 故障成因出口 / Fault cause outlet *)
    bError      : BOOL;                      (* 故障锁存标志 [-] / Fault latch flag *)
END_VAR
VAR
    _eState   : E_DL_FcqState := E_DL_FcqState.eIdle;     (* 内部相位（CASE 唯一写入目标） / Internal phase *)
    _eCause   : E_DL_FcqCause := E_DL_FcqCause.eNone;     (* 故障成因锁存量 / Latched cause *)
    rtReq     : R_TRIG;                     (* 申请沿实例，段 0 无条件调用 / Request edge *)
    rtDone    : R_TRIG;                     (* 完成沿实例，段 0 无条件调用 / Done edge *)
    rtReset   : R_TRIG;                     (* 复位沿实例，段 0 无条件调用 / Reset edge *)
    _anId     : ARRAY[1..8] OF INT;         (* 队列通道号槽 [—] / Queue id slots *)
    _anPrio   : ARRAY[1..8] OF INT;         (* 队列优先级槽 [-] / Queue priority slots *)
    _nDepth   : INT;                        (* 队列深度锁存 [条] / Depth latch *)
    _nDispId  : INT;                        (* 派发通道号锁存 [-] / Dispatch id latch *)
    _nPrioDispL : INT;                      (* 派发通道优先级锁存（抢占判据用）[-] / Dispatched prio latch *)
    _bDisp    : BOOL;                       (* 派发有效锁存 [-] / Dispatch valid latch *)
    _bPreempt : BOOL;                       (* 抢占单拍量 [-] / Preempt pulse work *)
    _bEvict   : BOOL;                       (* 摘除单拍量 [-] / Evict pulse work *)
    _bFull    : BOOL;                       (* 队满单拍量 [-] / Full pulse work *)
    _nSel     : INT;                        (* 最高优先级选中槽（每趟重算）[-] / Selected slot *)
    _i        : INT;                        (* 搬移游标（每趟重置，R227）[-] / Shift cursor *)
    _nDone    : UDINT;                      (* 收口计数锁存 [次] / Done count latch *)
    _bFault   : BOOL;                       (* 故障锁存位 / Latched fault bit *)
    _bCfgBad  : BOOL;                       (* 组态非法当拍量 / Illegal config this scan *)
END_VAR
VAR CONSTANT
    DL_FCQ_QMAX : INT := 8;                  (* 队列容量 [条] / Queue capacity *)
    DL_FCQ_IDMAX: INT := 99;                 (* 通道号上限 [-] / Channel id max *)
END_VAR

(* —— 段 0：当拍判据派生 + 沿实例无条件刷新（R228A） —— *)
_bCfgBad := (bReq AND ((nChanId < 1) OR (nChanId > DL_FCQ_IDMAX) OR (nPrio < 0) OR (nPrio > 3)));   (* 组态闸：申请沿域闸（R151） / Config gate on request domain *)
rtReq(CLK := bReq);                          (* 申请沿每拍必调 / Request edge every scan *)
rtDone(CLK := bChanDone);                    (* 完成沿每拍必调 / Done edge every scan *)
rtReset(CLK := bReset);                      (* 复位沿每拍必调 / Reset edge every scan *)

(* —— 段 1：单拍量预清零（R107） —— *)
_bPreempt := FALSE;                          (* 抢占脉冲预清，唯一分支置位 / Preempt preset *)
_bEvict := FALSE;                            (* 摘除脉冲预清 / Evict preset *)
_bFull := FALSE;                             (* 队满脉冲预清 / Full preset *)
_nSel := 0;                                  (* 选中槽预清（每趟重算，R285） / Selected slot preset *)

(* —— 段 2：复位沿处理（作用域：清故障 + 清队列 + 清派发 + 清计数 + 迁 eIdle，R283 逐项声明） —— *)
IF rtReset.Q THEN
    _bFault := FALSE;                        (* 清故障锁存 / Clear fault *)
    _eCause := E_DL_FcqCause.eNone;          (* 清成因 / Clear cause *)
    _nDepth := 0;                            (* 清队列深度 / Clear depth *)
    _nDispId := 0;                           (* 清派发号 / Clear dispatch id *)
    _nPrioDispL := 0;                        (* 清派发优先级锁存 / Clear prio latch *)
    _bDisp := FALSE;                         (* 清派发有效 / Clear valid *)
    nDispatchId := 0;                        (* 清派发出口 / Clear outlet *)
    _nDone := 0;                             (* 清收口计数 / Clear done count *)
    _eState := E_DL_FcqState.eIdle;          (* 迁待机相 / Back to idle *)
END_IF

(* —— 段 3：组态闸故障锁存（R45 配对；锁存至复位沿，R189） —— *)
IF _bCfgBad AND NOT _bFault THEN
    _bFault := TRUE;                         (* 锁存故障位 / Latch fault *)
    _eCause := E_DL_FcqCause.eCfgIllegal;    (* 成因：组态非法 / Cause: illegal config *)
    _eState := E_DL_FcqState.eFault;         (* 同步迁故障相 / Migrate to fault *)
END_IF

(* —— 段 4：CASE 主状态机（ELSE 兜底迁 eFault，红线 6） —— *)
CASE _eState OF
    E_DL_FcqState.eIdle:                     (* 待机相 / Idle *)
        IF bEnable AND NOT _bFault THEN
            _eState := E_DL_FcqState.eDispatch;   (* 进入调度 / Enter dispatch *)
        END_IF
    E_DL_FcqState.eDispatch:                 (* 调度相：入队 + 抢占 + 摘除 + 收口 + 派发 / Dispatch *)
        IF NOT bEnable THEN
            _eState := E_DL_FcqState.eIdle;  (* 失能回待机（派发保持，R191 声明） / Back to idle, dispatch held *)
        ELSE
            IF rtReq.Q THEN                  (* 申请沿：入队 / Enqueue on edge *)
                IF _nDepth < DL_FCQ_QMAX THEN
                    _nDepth := _nDepth + 1;  (* 深度 +1 / Depth up *)
                    _anId[_nDepth] := nChanId;       (* 尾插通道号 / Append id *)
                    _anPrio[_nDepth] := nPrio;       (* 尾插优先级 / Append prio *)
                ELSE
                    _bFull := TRUE;          (* 队满拒收单拍（不缓存，边界①） / Full reject *)
                END_IF
            END_IF
            IF _bDisp AND bChanFault THEN    (* 运行通道故障：摘除不回队 / Evict on fault *)
                _bEvict := TRUE;             (* 摘除单拍 / Evict pulse *)
                _bDisp := FALSE;             (* 撤派发 / Drop dispatch *)
            END_IF
            IF _bDisp AND rtDone.Q THEN      (* 正常收口 / Normal done *)
                _nDone := _nDone + 1;        (* 收口计数（UDINT 回绕 ≈ 49 天 @1kHz，工程安全） / Count done *)
                _bDisp := FALSE;             (* 撤派发 / Drop dispatch *)
            END_IF
            IF _bDisp AND rtReq.Q AND (NOT _bFull) AND (nPrio < _nPrioDispL) AND (_nDepth < DL_FCQ_QMAX) THEN
                (* 抢占：更优优先级申请且队列可容纳回队件 / Preempt: better prio + room for requeue *)
                _i := _nDepth;               (* 队列后移游标自尾起（R227） / Shift cursor from tail *)
                WHILE _i >= 1 DO             (* 全队后移一格腾出队头 / Shift back one slot *)
                    _anId[_i + 1] := _anId[_i];   (* 通道号后移 / Shift id *)
                    _anPrio[_i + 1] := _anPrio[_i];   (* 优先级后移 / Shift prio *)
                    _i := _i - 1;            (* 游标递退 / Cursor back *)
                END_WHILE
                _anId[1] := _nDispId;        (* 被抢占通道回队头 / Requeue preempted *)
                _anPrio[1] := 3;             (* 回队降为最低级（防反复抢占振荡，边界④） / Requeue at lowest prio *)
                _nDepth := _nDepth + 1;      (* 深度 +1 / Depth up *)
                _bPreempt := TRUE;           (* 抢占单拍 / Preempt pulse *)
                _bDisp := FALSE;             (* 撤当前派发 / Drop dispatch *)
            END_IF
            IF (NOT _bDisp) AND (_nDepth >= 1) THEN   (* 空派发且有队列：选最高优先级（数值最小，同级先入先出） / Pick best *)
                _nSel := 1;                  (* 先选队头（同级 FIFO 基准） / Seed with head *)
                _i := 2;                     (* 扫描游标重置（R227） / Scan cursor reset *)
                WHILE _i <= _nDepth DO       (* 逐槽找数值最小优先级 / Find min prio *)
                    IF _anPrio[_i] < _anPrio[_nSel] THEN
                        _nSel := _i;         (* 更优槽 / Better slot *)
                    END_IF
                    _i := _i + 1;            (* 游标递进 / Cursor advance *)
                END_WHILE
                _nDispId := _anId[_nSel];    (* 派发选中通道 / Dispatch selected *)
                _nPrioDispL := _anPrio[_nSel];   (* 锁存派发优先级（抢占判据基准） / Latch dispatched prio *)
                _bDisp := TRUE;              (* 置派发有效 / Set valid *)
                _i := _nSel;                 (* 删除搬移游标（R227） / Removal cursor *)
                WHILE _i < _nDepth DO        (* 后件前移补空 / Shift forward *)
                    _anId[_i] := _anId[_i + 1];   (* 通道号前移 / Shift id *)
                    _anPrio[_i] := _anPrio[_i + 1];   (* 优先级前移 / Shift prio *)
                    _i := _i + 1;            (* 游标递进 / Cursor advance *)
                END_WHILE
                _nDepth := _nDepth - 1;      (* 深度 -1 / Depth down *)
            END_IF
        END_IF
    E_DL_FcqState.eFault:                    (* 故障相：撤派发，仅复位沿出 / Fault *)
        _bDisp := FALSE;                     (* 故障相派发撤销（安全侧） / Drop dispatch in fault *)
        _nDispId := 0;                       (* 派发号清零 / Clear id *)
    ELSE                                     (* 非法相位兜底迁安全态 / Illegal phase fallback *)
        _eState := E_DL_FcqState.eFault;     (* 迁故障相 / To fault *)
        _bFault := TRUE;                     (* 同步锁存 / Latch *)
        _eCause := E_DL_FcqCause.ePhaseBad;  (* 成因：非法相位 / Cause: illegal phase *)
END_CASE

(* —— 段 5：出口映射（bError/eState 同源，R191） —— *)
nDispatchId := _nDispId;                     (* 派发号出口 / Dispatch id outlet *)
bDispatchValid := _bDisp;                    (* 派发有效出口 / Valid outlet *)
nQueueDepth := _nDepth;                      (* 深度出口 / Depth outlet *)
bQueueFull := _bFull;                        (* 队满脉冲出口 / Full outlet *)
bPreempt := _bPreempt;                       (* 抢占脉冲出口 / Preempt outlet *)
bEvict := _bEvict;                           (* 摘除脉冲出口 / Evict outlet *)
nDoneCnt := _nDone;                          (* 收口计数出口 / Done count outlet *)
bError := _bFault;                           (* 故障标志镜像 / Fault flag mirror *)
eState := _eState;                           (* 状态出口 / State outlet *)
eCause := _eCause;                           (* 成因出口 / Cause outlet *)
END_FUNCTION_BLOCK

(* ---- FB_DL_FormationTempRiseRate.st ---- *)
(*
  Component : FB_DL_FormationTempRiseRate
  Category  : DL_Process
  Type      : FB
  Version   : 1.0.0
  CodeSeg   : 16#06_0_3E
  Summary   : 化成温升速率监视与异常电芯截断：MA 前置平滑 + 速率微分 + 工艺窗分级报警 + 截断独立。
              Formation temp rise rate monitor: MA pre-smoothing plus rate differentiation, graded alarm, separate truncate.
  溯源声明  : 道莅自研 clean-room
  边界安全  : 温度非有限（NaN 自反 + Inf 上限）与负绝对温度域拦截；MA 点数域闸（2..16）；
              微分前置 MA 平滑防单拍毛刺误截断（按派单要点）；节拍正域闸与速率分母防除零；
              截断动作与报警分离，截断锁存仅手动复位沿可解除；TON/R_TRIG 每拍无条件刷新。
  复用      : 无
*)

FUNCTION_BLOCK FB_DL_FormationTempRiseRate
VAR_INPUT
    bRun        : BOOL;                 (* 监视使能 · Enable *)
    fTempC      : LREAL;                (* 电芯温度 [degC] · Cell temperature *)
    tPaceMs     : TIME  := T#1000MS;    (* 速率采样节拍 [ms] · Rate sample pace *)
    nMaPts      : INT   := 8;           (* MA 平滑点数 [点]，域 2 到 16 · MA smoothing points *)
    fRateHiKps  : LREAL := 0.5;         (* 高速升率报警阈 [K/s] · High rise rate threshold *)
    fRateCritKps: LREAL := 1.0;         (* 临界升率截断阈 [K/s] · Critical truncate threshold *)
    bTruncReset : BOOL;                 (* 截断手动复位 [事件]，沿触发 · Truncate manual reset *)
    fEps        : LREAL := 1.0E-6;      (* 浮点判零容差 [实数域] · Floating zero tolerance *)
END_VAR
VAR_OUTPUT
    fMaTempC  : LREAL;                  (* 平滑后温度 [degC] · Smoothed temperature *)
    fRateKps  : LREAL;                  (* 温升速率 [K/s] · Temperature rise rate *)
    bWarnHi   : BOOL;                   (* 高速升率报警（非锁存）· High rate warning *)
    bTruncate : BOOL;                   (* 异常截断指令锁存 · Latched truncate command *)
    bError    : BOOL;                   (* 故障标志，与故障码配对 · Fault flag paired with codes *)
    uErrorId  : UDINT;                  (* 事件码 16#0000_003E，0 无事件 · Event code *)
END_VAR
VAR
    uCode   : WORD;     (* 码位暂存，每拍重算 [码] · Code staging *)
    tonPace : TON;      (* 采样节拍 [ms]，自复位振荡 · Sample pace timer, self-reset *)
    rTrigRst: R_TRIG;   (* 截断复位沿检测 · Truncate reset edge *)
    aRing   : ARRAY[1..16] OF LREAL;    (* 温度环形缓冲 [degC] · Temperature ring buffer *)
    nHead   : INT;      (* 环形头下标 [索引] · Ring head index *)
    nFill   : INT;      (* 已填充点数 [点] · Filled point count *)
    fMaPrv  : LREAL;    (* 上节拍平滑温度快照 [degC] · Previous MA snapshot *)
    fDtS    : LREAL;    (* 节拍秒值 [s]，一次导出 · Pace seconds *)
    bSnapOk : BOOL;     (* 快照有效标志 · Snapshot validity *)
    bSigOk  : BOOL;     (* 输入有效标志 · Input validity flag *)
    bTick   : BOOL;     (* 采样到点脉冲 [脉冲] · Sample tick pulse *)
    nI      : INT;      (* 求和循环下标 [索引] · Sum loop index *)
    nCycles : UDINT;    (* 有效采样拍计数 [拍]，防回卷 · Sample count *)
END_VAR
VAR CONSTANT
    DL_FTR_ABS0 : LREAL := 273.15;      (* 绝对零度 [degC] · Absolute zero *)
    DL_FTR_NMAX : INT := 16;            (* 环形容量 [点] · Ring capacity *)
    DL_FTR_WRAP : UDINT := 4294967290;  (* 计数防回卷余量 [拍] · Counter wrap guard *)
END_VAR

(* === 段 0 · 实例刷新（每拍无条件，红线 7）=== *)
tonPace(IN := NOT tonPace.Q, PT := tPaceMs);    (* 节拍自复位振荡 / Self-reset pace *)
rTrigRst(CLK := bTruncReset);                   (* 截断复位沿 / Truncate reset edge *)
bTick := tonPace.Q;                             (* 采样脉冲 / Sample tick *)

(* === 段 1 · 输入校验与量程闸 === *)
uCode := 16#0000;                       // 每拍清码（可达清零基线）/ Clear codes each scan
bSigOk := (fTempC = fTempC) AND (ABS(fTempC) < 1.0E308)             // 非有限拦截 / Non-finite guard
          AND (fTempC > -DL_FTR_ABS0 + fEps)                         // 绝对零物理域闸 / Physical domain
          AND (nMaPts >= 2) AND (nMaPts <= DL_FTR_NMAX)              // MA 点数域闸 / MA point gate
          AND (tPaceMs > T#0MS)                                      // 节拍正域闸 / Pace gate
          AND (fRateHiKps > 0.0) AND (fRateCritKps > fRateHiKps);    // 阈值序闸 / Threshold order gate
IF fDtS < fEps THEN
    fDtS := DINT_TO_LREAL(TIME_TO_DINT(tPaceMs)) / 1000.0;      (* 节拍秒值一次导出 / Derive once *)
END_IF
IF NOT bSigOk THEN
    uCode := 16#003E;                   // 故障级：域外，监视冻结 / Fault: domain invalid
END_IF

(* === 段 2 · 主逻辑：MA 平滑与速率微分 === *)
IF bSigOk THEN
    IF bTick THEN
        IF nHead < 1 THEN
            nHead := 1;                 (* 头下标初值钳 1，防零下标越界 / Clamp the head to one *)
        END_IF
        IF nFill < nMaPts THEN
            nFill := nFill + 1;         (* 未满先增填充 / Grow fill *)
        END_IF
        aRing[nHead] := fTempC;         (* 写入采样 / Write the sample *)
        nHead := (nHead MOD DL_FTR_NMAX) + 1;   (* 头下标循环推进 / Advance the head *)
        fMaTempC := 0.0;                (* 平滑和清零 / Clear the sum *)
        FOR nI := 1 TO nMaPts DO
            IF nI <= nFill THEN
                fMaTempC := fMaTempC + aRing[nI];   (* 窗内累加 / Accumulate in window *)
            END_IF
        END_FOR
        fMaTempC := fMaTempC / UDINT_TO_LREAL(INT_TO_UDINT(nFill));     (* MA 均值 [degC] / MA mean *)
        IF bSnapOk THEN
            fRateKps := (fMaTempC - fMaPrv) / fDtS;     (* 速率微分 [K/s]，MA 前置平滑 / Differentiated rate *)
            IF fRateKps < 0.0 THEN
                fRateKps := 0.0;        (* 降温段速率钳零 / Clamp negative rate *)
            END_IF
        END_IF
        fMaPrv := fMaTempC;             (* 快照更新 / Update the snapshot *)
        bSnapOk := TRUE;                (* 快照有效 / Snapshot valid *)
        IF nCycles < DL_FTR_WRAP THEN
            nCycles := nCycles + 1;     (* 有效采样计数 / Count samples *)
        END_IF
    END_IF
    bWarnHi := (fRateKps > fRateHiKps); (* 高速升率报警（非锁存自清）/ Non-latched warning *)
    IF fRateKps > fRateCritKps THEN
        bTruncate := TRUE;              (* 临界截断锁存 / Latch the truncate *)
    END_IF
END_IF

(* === 段 3 · 输出映射与故障码 === *)
IF rTrigRst.Q THEN
    bTruncate := FALSE;                 (* 截断仅手动复位沿可解除（可达路径）/ Manual reset clears truncate *)
END_IF
IF NOT bRun THEN
    bWarnHi := FALSE;                   (* 撤使能报警清零 / Clear warnings on disable *)
END_IF
bError := (uCode <> 16#0000);           (* 故障标志配对 / Fault flag paired *)
uErrorId := WORD_TO_UDINT(uCode);       (* 码位单点写入（16#0000_003E 形态）/ Single write point *)
END_FUNCTION_BLOCK
